(* IEC 61131-3 sources: daoli-st-library/DL_Process (part 21) *)

(* ---- FB_DL_AnnealCoolRateCtrl.st ---- *)
(*
  Name: FB_DL_AnnealCoolRateCtrl
  Category: DL_Process
  Version: 1.0.0
  Round: R89 / 2026-11-25
  开源溯源：clean-room 自研（族 锻造加热退火，ST 开源生态实测 0 命中，无外部代码引入）
  功能：退火冷却速率控制：微分实测降温速率，超速报警；同时做超温（实测高于设定 + 容差）保护。
  边界条件：① 四浮点入参全部过非有限闸；配置越域或失能进冻结分支：输出保持末值 + xValid = FALSE（R191）；
            ② 归因分离（R190）：超速与超温各有独立内部成员 _bOverRate / _bOverTemp，出口合并为 xRateAlarm，
               两成因赋值点互不共用，头注释声明合并口径；
            ③ 微分为一阶差分：速率 = (上拍温度 − 本拍温度)/周期 × 60，正值为降温方向 [℃/min]；
            ④ 首扫 _bInit 以当前温度播种上拍快照，避免首拍出现虚假大速率；非法周期取 10 ms 缺省。
  量纲自证：℃ ÷ s × 60 = ℃/min；容差 ℃ 与温度同量纲。
*)
FUNCTION_BLOCK FB_DL_AnnealCoolRateCtrl
VAR_INPUT
    xEnable : BOOL;             (* 使能 [-] Enable *)
    fTempActC : REAL;           (* 炉温实测 [℃] Furnace temperature actual [degC] *)
    fTempSpC : REAL;            (* 炉温设定 [℃] Furnace temperature setpoint [degC] *)
    fCoolRateMaxCpm : REAL;     (* 最大允许降温速率 [℃/min] Maximum allowed cooling rate [degC/min] *)
    fCycleS : REAL;             (* 扫描周期 [s] Scan cycle [s] *)
END_VAR
VAR_OUTPUT
    fRateActCpm : REAL;         (* 实测降温速率（正值为降温） [℃/min] Actual cooling rate [degC/min] *)
    xRateAlarm : BOOL;          (* 超速或超温报警（归因见内部成员） [-] Over-rate or over-temperature alarm *)
    xValid : BOOL;              (* 配置与链路有效 [-] Configuration and chain valid *)
END_VAR
VAR
    _bInit : BOOL := FALSE;     (* 首扫初始化标志 [-] First-scan init flag *)
    _bCfgBad : BOOL := FALSE;   (* 配置非法当拍量 [-] Configuration bad *)
    _bCalcOk : BOOL := FALSE;   (* 本拍计算有效 [-] Calculation valid this scan *)
    _bOverRate : BOOL := FALSE; (* 超速成因（独立成员） [-] Over-rate cause *)
    _bOverTemp : BOOL := FALSE; (* 超温成因（独立成员） [-] Over-temperature cause *)
    _fPrev : REAL := 0.0;       (* 上拍温度快照（首扫播种） [℃] Previous temperature snapshot [degC] *)
    _fRate : REAL := 0.0;       (* 速率保持量 [℃/min] Rate hold [degC/min] *)
    _fCy : REAL := 0.01;        (* 当拍有效周期 [s] Effective cycle [s] *)
END_VAR
VAR CONSTANT
    DL_ACRC_EPS : REAL := 1.0E-9;       (* 判据容差 [-] Criterion tolerance *)
    DL_ACRC_CYDEF : REAL := 0.01;       (* 缺省扫描周期 [s] Default scan cycle [s] *)
    DL_ACRC_SECMIN : REAL := 60.0;      (* 每秒 → 每分钟换算 [s/min] Second to minute *)
    DL_ACRC_TOL : REAL := 5.0;          (* 超温容差 [℃] Over-temperature tolerance [degC] *)
    DL_ACRC_TMIN : REAL := 0.0;         (* 温度下限 [℃] Temperature floor [degC] *)
    DL_ACRC_TMAX : REAL := 1400.0;      (* 温度上限 [℃] Temperature ceiling [degC] *)
    DL_ACRC_RMIN : REAL := 0.1;         (* 允许速率下限 [℃/min] Rate floor [degC/min] *)
    DL_ACRC_RMAX : REAL := 100.0;       (* 允许速率上限 [℃/min] Rate ceiling [degC/min] *)
END_VAR
(* 首扫初始化：以当前温度播种上拍快照，避免虚假大速率（R310） *)
IF NOT _bInit THEN
    _fPrev := fTempActC;
    _fRate := 0.0;
    _bInit := TRUE;
END_IF
(* 周期派生：非法周期取 10 ms 缺省（步长不塌零，除零结构性排除） *)
IF (fCycleS > 0.0) AND (fCycleS <= 1.0) THEN
    _fCy := fCycleS;
ELSE
    _fCy := DL_ACRC_CYDEF;
END_IF
(* 非有限闸（NaN 自反 + Inf 差值自减）+ 组态域闸：四浮点入参全枚举（R272） *)
_bCfgBad := (fTempActC <> fTempActC) OR ((fTempActC - fTempActC) <> 0.0)
         OR (fTempSpC <> fTempSpC) OR ((fTempSpC - fTempSpC) <> 0.0)
         OR (fCoolRateMaxCpm <> fCoolRateMaxCpm) OR ((fCoolRateMaxCpm - fCoolRateMaxCpm) <> 0.0)
         OR (fCycleS <> fCycleS) OR ((fCycleS - fCycleS) <> 0.0)
         OR (fTempActC < DL_ACRC_TMIN) OR (fTempActC > DL_ACRC_TMAX)
         OR (fTempSpC < DL_ACRC_TMIN) OR (fTempSpC > DL_ACRC_TMAX)
         OR (fCoolRateMaxCpm < DL_ACRC_RMIN) OR (fCoolRateMaxCpm > DL_ACRC_RMAX);
_bCalcOk := xEnable AND (NOT _bCfgBad);
IF _bCalcOk THEN
    (* 一阶差分：正值为降温方向，量纲 ℃/s × 60 = ℃/min *)
    _fRate := ((_fPrev - fTempActC) / _fCy) * DL_ACRC_SECMIN;
    (* 归因分离：超速与超温各写各的成员，互不共用赋值点（R190） *)
    _bOverRate := _fRate > fCoolRateMaxCpm;
    _bOverTemp := fTempActC > (fTempSpC + DL_ACRC_TOL);
    (* 快照推进放在有效计算之后，冻结时快照不动 *)
    _fPrev := fTempActC;
ELSE
    _bOverRate := FALSE;
    _bOverTemp := FALSE;
    _fPrev := fTempActC;                    (* 冻结拍也同步快照，恢复时不产生阶跃虚假速率 *)
END_IF
(* 统一出口（单点赋值）：冻结分支保持末次有效速率，保持量为已过闸的有限值（R273） *)
fRateActCpm := _fRate;
xRateAlarm := (_bOverRate OR _bOverTemp) AND _bCalcOk;
xValid := _bCalcOk;
END_FUNCTION_BLOCK

(* ---- FB_DL_BacdHvacPoll.st ---- *)
(*
  ==================================================================
  组件名 Component  : FB_DL_BacdHvacPoll
  分类   Category   : DL_Process
  版本   Version    : 1.0.1
  功能   Purpose    : BA 顺控 BACnet / Modbus 轮询行。按固定轮询间隔对 1..16 台现场
                      设备做轮询：发出轮询触发后等响应超时窗，收到响应即置在线位并
                      清重试计数；超时即重试，重试次数用尽置离线位。每轮完成后索引
                      前进并跳过离线设备（全部离线时仍逐台尝试以探测恢复），并输出
                      在线 / 离线掩码字、轮询计数与超时计数。
  溯源   Origin     : BACnet / Modbus 轮询调度为公开现场总线通信语义；本件为 clean-room
                      实现，仅借鉴来源分类与参数域组织（来源标签 roadmap-p2-bacd），
                      道莅原创设计，未复制任何闭源代码行。
  平台   Platform   : 纯 IEC 61131-3（TON / R_TRIG / WORD / SHL，无私有库）
  作者   Author     : 道莅代码库 · PLC 编程专家（R55）
  ------------------------------------------------------------------
  同拍双窗配比约束（R100）：tRespTo 必须小于 tPollInt —— 响应超时窗短于轮询间隔窗，
                      两窗职责分离：tPollInt 定节拍，tRespTo 判单台失败；超时窗覆盖整个
                      间隔会使下一拍无法发出轮询，配比反置在组态域闸内直接判故障。
  边界 Boundary     :
                      一 本件只出轮询触发与在线掩码，不做协议编解码、不写设备（属主边界）；
                      二 轮询间隔用自复位周期 TON（周期脉冲发生器用法，R328 适用方向）；
                      三 响应超时件 IN 串「等待响应相」闸与「响应已到」补集，不跨相累计；
                      四 设备索引一律回钳 1..16，跳过离线设备的循环有守护上限防死循环；
                      五 无全局变量、无外部变量声明、无物理地址寻址；
                      六 eNoDevice 为预留恒空成员：设备数为零已由组态域闸判
                         eCfgIllegal（故障级），信息级 eNoDevice 不可达，保留成员
                         以稳定接口（R56 返修留痕）。
  输出契约 Output contract:
                      nPollIdx 为当前轮询设备号（1..nDevCount），无设备时保持 1；
                      wOnlineMask / wOfflineMask 位 i-1 对应设备 i，
                      自证向量：仅 1 号设备离线 → 16#0001，仅 16 号设备离线 → 16#8000；
                      bPollTrig 与 bRespTimeout 各为单拍脉冲（内部位置位、出口映射后撤销）；
                      eCause 故障级成因与 bError 配对（R45），信息级永不置 bError。
  修订记录 Revision  :
    2026-11-20  v1.0.0  R55 首版（批 4 · 序号 20）
    2026-11-20  v1.0.1  R56 返修（7.1）：段 7 删除恒假死分支（判量 _nUseCount 经段 3
                        回钳恒 ≥1，信息级 eNoDevice 不可达），「设备数为零」语义改由
                        组态域闸 eCfgIllegal（故障级）承载；_nCurRetry 声明经核验
                        已在 VAR 区在位（7 处引用合法）。
  ==================================================================
*)

TYPE E_DL_BhdPhase :
(
    eIdle  := 0,        // 空闲：未使能或已停轮询 / idle, disabled or polling stopped
    ePoll  := 10,       // 发出：本拍发出轮询触发 / issuing, the poll trigger is raised this scan
    eWait  := 20,       // 等响应：等响应或超时 / waiting, for the response or the timeout
    eFault := 90        // 故障：组态非法锁存 / fault, illegal configuration latched
);
END_TYPE

TYPE E_DL_BhdCause :
(
    eNone       := 0,   // 无成因 / no cause
    eCfgIllegal := 1,   // 组态非法：设备数、重试上限或时间引脚越域（故障级，与 bError 配对）/ illegal config, device count, retry cap or time pin out of domain
    eDevOffline := 2,   // 有设备重试用尽转离线（信息级）/ a device exhausted its retries and went offline, informational
    eAllOffline := 3,   // 全部设备离线，仍逐台尝试探测恢复（信息级）/ every device is offline and the scan still probes for recovery
    eNoDevice   := 4    // 设备数为零（预留恒空，语义由 eCfgIllegal 承载，R56 留痕）/ no device configured, reserved always empty, carried by eCfgIllegal
);
END_TYPE

FUNCTION_BLOCK FB_DL_BacdHvacPoll
VAR_INPUT
    bEnable     : BOOL := TRUE;              // 使能，失能时停轮询并保持掩码 [-] / enable, polling stops and the masks hold when disabled
    bReset      : BOOL := FALSE;            // 复位上升沿清故障锁存、掩码与重试 [-] / reset rising edge clears the fault latch, the masks and the retries
    nDevCount   : INT := 8;                  // 轮询设备数 [台]，域 1..16 / polled device count [unit], domain 1 to 16
    nRetryMax   : INT := 2;                  // 单设备重试上限 [次]，域 0..9 / per device retry ceiling [count], domain 0 to 9
    tPollInt    : TIME := T#1S;              // 轮询间隔 [毫秒]，域 大于零 / poll interval [millisecond], domain above zero
    tRespTo     : TIME := T#500MS;           // 响应超时 [毫秒]，域 大于零 / response timeout [millisecond], domain above zero
    bRespPulse  : BOOL := FALSE;             // 响应到达脉冲（对应当前轮询设备）[-] / response arrival pulse for the currently polled device
END_VAR
VAR_OUTPUT
    nPollIdx    : INT := 1;                  // 当前轮询设备号 [设备号] / currently polled device number
    bPollTrig   : BOOL := FALSE;             // 轮询触发单拍脉冲 [-] / poll trigger single-shot pulse
    bRespTimeout: BOOL := FALSE;             // 响应超时单拍脉冲 [-] / response timeout single-shot pulse
    wOnlineMask : WORD := 16#0000;           // 在线设备掩码，位 i-1 对应设备 i [-] / online device mask, bit i minus one maps to device i
    wOfflineMask: WORD := 16#0000;           // 离线设备掩码，位 i-1 对应设备 i [-] / offline device mask, bit i minus one maps to device i
    uPollCnt    : UDINT := 0;                // 累计轮询次数（饱和到上限）[次] / total poll count, saturated [count]
    uTimeoutCnt : UDINT := 0;                // 累计响应超时次数（饱和到上限）[次] / total response timeout count, saturated [count]
    nOfflineCnt : INT := 0;                  // 当前离线设备数 [台] / current offline device count [unit]
    nCurRetry   : INT := 0;                  // 当前设备已重试次数 [次] / retries already spent on the current device [count]
    ePhase      : E_DL_BhdPhase := E_DL_BhdPhase.eIdle; // 相位出口 [枚举] / phase outlet [enum]
    eCause      : E_DL_BhdCause := E_DL_BhdCause.eNone; // 成因出口 [枚举] / cause outlet [enum]
    bError      : BOOL := FALSE;             // 故障锁存标志 [-] / fault latch flag
END_VAR
VAR
    rtResp      : R_TRIG;                    // 响应沿检测，段 0 无条件刷新 / response edge detector, refreshed unconditionally in segment zero
    rtReset     : R_TRIG;                    // 复位沿检测，段 0 无条件刷新 / reset edge detector, refreshed unconditionally in segment zero
    tonPollInt  : TON;                       // 轮询间隔周期计时（自复位式）/ poll interval timer, self resetting
    tonResp     : TON;                       // 响应超时计时，段 0 无条件刷新 / response timeout timer, refreshed unconditionally in segment zero
    _ePhase     : E_DL_BhdPhase := E_DL_BhdPhase.eIdle;   // 内部相位，CASE 唯一写入目标 / internal phase, the only CASE write target
    _eCause     : E_DL_BhdCause := E_DL_BhdCause.eNone;   // 信息级成因，每拍重算 / informational cause, recomputed every scan
    _eFaultCause: E_DL_BhdCause := E_DL_BhdCause.eNone;   // 故障级成因，锁存至复位沿 / fault cause, latched until the reset edge
    _bFault     : BOOL := FALSE;             // 故障锁存位 [-] / fault latch bit
    _bInit      : BOOL := FALSE;             // 首扫初始化完成标志（R310）/ first scan initialisation flag
    _bCfgBad    : BOOL := FALSE;             // 组态非法判定 [-] / illegal configuration verdict
    _bPollInt   : BOOL := FALSE;             // 轮询触发内部位，统一出口映射 / internal poll trigger bit, mapped at the unified outlet
    _bToInt     : BOOL := FALSE;             // 超时脉冲内部位，统一出口映射 / internal timeout bit, mapped at the unified outlet
    _bOfflineNew: BOOL := FALSE;             // 本拍有新设备转离线 [-] / a device went offline this scan
    _bAllOff    : BOOL := FALSE;             // 全部设备离线 [-] / every device is offline
    _bFound     : BOOL := FALSE;             // 跳过循环命中标志 [-] / hit flag of the skip loop
    _bIsOffline : BOOL := FALSE;             // 被检设备是否离线 [-] / whether the checked device is offline
    _nUseCount  : INT := 1;                  // 钳定后的设备数 [台] / clamped device count [unit]
    _nRetryUse  : INT := 1;                  // 钳定后的重试上限 [次] / clamped retry ceiling [count]
    _nIdx       : INT := 1;                  // 设备索引（回钳 1..16）[设备号] / device index clamped one through sixteen
    _nGuard     : INT := 0;                  // 跳过循环守护计数 [次] / skip loop guard [count]
    _nIdxProbe  : INT := 1;                  // 离线统计探测索引 [设备号] / probe index for the offline statistics
    _nCurRetry  : INT := 0;                  // 当前设备重试计数（声明补齐，R55 终审）/ current device retry counter, declaration completed at R55 review
    _nOfflineCnt: INT := 0;                  // 本轮统计离线设备数工作值（出口映射源）[台] / offline device count working value, source of the outlet [unit]
    _wOff       : WORD := 16#0000;           // 离线掩码工作字 / offline mask working word
    _wOn        : WORD := 16#0000;           // 在线掩码工作字（按位或累计）/ online mask working word
    _wBit       : WORD := 16#0001;           // 本设备位掩码，先移位后置位（R327）/ device bit mask, shift before setting
    _uPoll      : UDINT := 0;                // 轮询计数工作值 [次] / poll count working value [count]
    _uTo        : UDINT := 0;                // 超时计数工作值 [次] / timeout count working value [count]
END_VAR
VAR CONSTANT
    DL_BHD_MAX      : INT := 16;             // 设备容量与索引回钳上界 [台] / device capacity and index clamp upper bound
    DL_BHD_RETRY_MAX: INT := 9;              // 重试上限的钳定上限 [次] / clamp ceiling of the retry cap [count]
    DL_BHD_CNT_MAX  : UDINT := 2000000000;   // 计数饱和上限（常量在 DINT 可表范围内）[次] / count saturation ceiling, the constant fits in DINT
    DL_BHD_MASK_NONE: WORD := 16#0000;       // 空掩码常量 [-] / empty mask constant
    DL_BHD_MASK_ONE : WORD := 16#0001;       // 单位位常量 [-] / single bit constant
END_VAR

// 段 0｜定时器与沿检测无条件周期刷新（禁入分支）；轮询间隔用自复位式周期发生器 / segment 0, unconditional refresh with a self resetting periodic generator
rtResp(CLK := bRespPulse); // 响应沿无条件刷新 / unconditional refresh of the response edge
rtReset(CLK := bReset); // 复位沿无条件刷新 / unconditional refresh of the reset edge
tonPollInt(IN := (NOT tonPollInt.Q) AND bEnable AND (NOT _bFault), PT := tPollInt); // 轮询间隔周期发生器，Q 到时下一拍即重启（R328 周期脉冲方向）/ periodic poll generator that restarts right after its own pulse
tonResp(IN := (_ePhase = E_DL_BhdPhase.eWait) AND (NOT rtResp.Q) AND (NOT _bFault), PT := tRespTo); // 响应超时，IN 串等待相闸与响应到达补集 / response timeout with the waiting gate and the response complement on IN

// 段 1｜首扫初始化（R310）/ segment 1, first scan initialisation
IF NOT _bInit THEN // 首扫一拍 / the very first scan
    _bInit := TRUE; // 置首扫完成标志 / raise the first scan flag
    _ePhase := E_DL_BhdPhase.eIdle; // 相位从空闲起步 / the phase starts from idle
    _eCause := E_DL_BhdCause.eNone; // 信息级成因清零 / clear the informational cause
    _eFaultCause := E_DL_BhdCause.eNone; // 故障级成因清零 / clear the fault cause
    _bFault := FALSE; // 故障锁存清零 / clear the fault latch
    _wOff := DL_BHD_MASK_NONE; // 离线掩码清零 / clear the offline mask
    _wOn := DL_BHD_MASK_NONE; // 在线掩码清零 / clear the online mask
    _nIdx := 1; // 索引归位 / park the index at one
    _uPoll := 0; // 轮询计数清零 / clear the poll count
    _uTo := 0; // 超时计数清零 / clear the timeout count
END_IF

// 段 2｜复位沿作用域：清锁存 / 清掩码 / 清计数与索引（四项逐项声明）/ segment 2, reset edge scope declared item by item
IF rtReset.Q THEN // 复位沿 / reset edge
    _bFault := FALSE; // 作用域一：清故障锁存 / scope one, clear the fault latch
    _eFaultCause := E_DL_BhdCause.eNone; // 作用域一：清故障级成因 / scope one, clear the fault cause
    _wOff := DL_BHD_MASK_NONE; // 作用域二：清离线掩码 / scope two, clear the offline mask
    _wOn := DL_BHD_MASK_NONE; // 作用域二：清在线掩码 / scope two, clear the online mask
    _nIdx := 1; // 作用域三：索引归位 / scope three, park the index
    _nCurRetry := 0; // 作用域三：清重试计数 / scope three, clear the retry count
    _ePhase := E_DL_BhdPhase.eIdle; // 作用域四：迁回空闲相 / scope four, migrate back to idle
    _bPollInt := FALSE; // 作用域四：清轮询脉冲内部位 / scope four, clear the internal poll bit
    _bToInt := FALSE; // 作用域四：清超时脉冲内部位 / scope four, clear the internal timeout bit
END_IF

// 段 3｜组态域闸（R151 全覆盖）/ segment 3, configuration domain gate over every pin
_bCfgBad := FALSE; // 组态非法预置假 / preset the illegal configuration verdict to false
IF (nDevCount < 1) OR (nDevCount > DL_BHD_MAX) THEN // 设备数越域 / the device count is out of domain
    _bCfgBad := TRUE; // 判非法 / mark illegal
END_IF
IF (nRetryMax < 0) OR (nRetryMax > DL_BHD_RETRY_MAX) THEN // 重试上限越域 / the retry cap is out of domain
    _bCfgBad := TRUE; // 判非法 / mark illegal
END_IF
IF (tPollInt <= T#0S) OR (tRespTo <= T#0S) THEN // 时间引脚非正 / a time pin is not positive
    _bCfgBad := TRUE; // 判非法 / mark illegal
END_IF
IF tRespTo >= tPollInt THEN // 响应超时窗不得覆盖整个轮询间隔（配比约束，R100）/ the response window must not swallow the whole poll interval
    _bCfgBad := TRUE; // 判非法 / mark illegal
END_IF
IF _bCfgBad AND (NOT _bFault) THEN // 组态非法且未锁存 / illegal configuration and not yet latched
    _bFault := TRUE; // 置故障锁存 / raise the fault latch
    _eFaultCause := E_DL_BhdCause.eCfgIllegal; // 故障级成因 (R45 配对 bError) / fault grade cause paired with bError
    _ePhase := E_DL_BhdPhase.eFault; // 迁故障相 / migrate to the fault phase
END_IF
_nUseCount := nDevCount; // 设备数直通 / the device count passes through
IF _nUseCount < 1 THEN // 下越界 / below the lower bound
    _nUseCount := 1; // 回钳到 1 / clamp to one
ELSIF _nUseCount > DL_BHD_MAX THEN // 上越界 / above the upper bound
    _nUseCount := DL_BHD_MAX; // 回钳到 16 / clamp to sixteen
END_IF
_nRetryUse := nRetryMax; // 重试上限直通 / the retry cap passes through
IF _nRetryUse < 0 THEN // 下越界（防御）/ below the lower bound as a defence
    _nRetryUse := 0; // 回钳到 0 / clamp to zero
ELSIF _nRetryUse > DL_BHD_RETRY_MAX THEN // 上越界 / above the upper bound
    _nRetryUse := DL_BHD_RETRY_MAX; // 回钳到 9 / clamp to nine
END_IF
IF _nIdx < 1 THEN // 索引下越界 / the index is below the lower bound
    _nIdx := 1; // 回钳到 1 / clamp to one
ELSIF _nIdx > _nUseCount THEN // 索引上越界 / the index is above the upper bound
    _nIdx := _nUseCount; // 回钳到末台 / clamp to the last unit
END_IF

// 段 4｜失效使能与设备位更新 / segment 4, enable handling and device bit updates
_eCause := E_DL_BhdCause.eNone; // 信息级成因每拍重算 / the informational cause is recomputed every scan
_bOfflineNew := FALSE; // 新转离线标志预置假 / preset the new offline flag to false
_bAllOff := FALSE; // 全离线标志每拍重算 / the all offline flag is recomputed every scan
IF NOT bEnable THEN // 失能：停轮询并保持掩码（R191 显式声明）/ disabled, polling stops and the masks hold
    _ePhase := E_DL_BhdPhase.eIdle; // 回空闲相 / return to idle
    _bPollInt := FALSE; // 撤轮询脉冲内部位 / withdraw the internal poll bit
    _bToInt := FALSE; // 撤超时脉冲内部位 / withdraw the internal timeout bit
END_IF
_wBit := SHL(DL_BHD_MASK_ONE, _nIdx - 1); // 当前设备位掩码，位移量 0..15 由索引回钳与容量常量证明 / the current device bit mask, the shift zero through fifteen is proven by the index clamp and the capacity constant
IF rtResp.Q AND (_ePhase = E_DL_BhdPhase.eWait) THEN // 等待相收到响应 / a response arrived while waiting
    _wOff := _wOff AND NOT _wBit; // 清离线位 / clear the offline bit
    _wOn := _wOn OR _wBit; // 置在线位 / set the online bit
    _nCurRetry := 0; // 清重试计数 / clear the retry count
    _ePhase := E_DL_BhdPhase.ePoll; // 本轮结束，转下一轮发出相 / the round is finished and the next issuing phase follows
    _bFound := FALSE; // 跳过命中标志预置假 / preset the skip hit flag to false
    _nGuard := 0; // 守护计数清零 / reset the guard
    WHILE (_nGuard < DL_BHD_MAX) AND (NOT _bFound) DO // 跳过离线设备，守护上限为容量 / skip offline devices with the capacity as the guard
        _nGuard := _nGuard + 1; // 守护计数递增 / increment the guard
        _nIdx := _nIdx + 1; // 索引前进 / advance the index
        IF _nIdx > _nUseCount THEN // 越过末台 / past the last unit
            _nIdx := 1; // 回卷到首台 / wrap back to the first unit
        END_IF
        _wBit := SHL(DL_BHD_MASK_ONE, _nIdx - 1); // 候选设备位掩码 / the candidate device bit mask
        _bIsOffline := ((_wOff AND _wBit) <> DL_BHD_MASK_NONE); // 候选设备是否离线 / whether the candidate is offline
        IF NOT _bIsOffline THEN // 候选在线 / the candidate is online
            _bFound := TRUE; // 命中 / hit
        END_IF
    END_WHILE
    IF NOT _bFound THEN // 全部离线，仍逐台尝试（探测恢复）/ every device is offline and probing continues
        _nIdx := _nIdx + 1; // 索引照常前进 / the index advances anyway
        IF _nIdx > _nUseCount THEN // 越过末台 / past the last unit
            _nIdx := 1; // 回卷到首台 / wrap back to the first unit
        END_IF
        _bAllOff := TRUE; // 置全离线标志 / raise the all offline flag
    END_IF
END_IF
IF tonResp.Q AND (_ePhase = E_DL_BhdPhase.eWait) THEN // 等待相超时 / the waiting phase timed out
    _bToInt := TRUE; // 超时脉冲内部位置位（统一出口映射，R187）/ raise the internal timeout bit, mapped at the unified outlet
    IF _uTo < DL_BHD_CNT_MAX THEN // 未达饱和上限 / below the ceiling
        _uTo := _uTo + 1; // 超时计数递增 / increment the timeout count
    END_IF
    IF _nCurRetry < _nRetryUse THEN // 重试未用尽 / retries remain
        _nCurRetry := _nCurRetry + 1; // 重试计数递增并立即重发 / increment the retry count and re-issue at once
        _ePhase := E_DL_BhdPhase.ePoll; // 回发出相重试同一台 / back to the issuing phase for the same unit
    ELSE // 重试用尽 / retries exhausted
        _wOff := _wOff OR _wBit; // 置离线位 / set the offline bit
        _wOn := _wOn AND NOT _wBit; // 清在线位 / clear the online bit
        _bOfflineNew := TRUE; // 记新转离线 / record the new offline event
        _nCurRetry := 0; // 重试计数清零 / clear the retry count
        _ePhase := E_DL_BhdPhase.ePoll; // 回发出相转下一台 / back to the issuing phase for the next unit
        _bFound := FALSE; // 跳过命中标志预置假 / preset the skip hit flag to false
        _nGuard := 0; // 守护计数清零 / reset the guard
        WHILE (_nGuard < DL_BHD_MAX) AND (NOT _bFound) DO // 跳过离线设备 / skip offline devices
            _nGuard := _nGuard + 1; // 守护计数递增 / increment the guard
            _nIdx := _nIdx + 1; // 索引前进 / advance the index
            IF _nIdx > _nUseCount THEN // 越过末台 / past the last unit
                _nIdx := 1; // 回卷到首台 / wrap back to the first unit
            END_IF
            _wBit := SHL(DL_BHD_MASK_ONE, _nIdx - 1); // 候选设备位掩码 / the candidate device bit mask
            _bIsOffline := ((_wOff AND _wBit) <> DL_BHD_MASK_NONE); // 候选设备是否离线 / whether the candidate is offline
            IF NOT _bIsOffline THEN // 候选在线 / the candidate is online
                _bFound := TRUE; // 命中 / hit
            END_IF
        END_WHILE
        IF NOT _bFound THEN // 全部离线 / every device is offline
            _bAllOff := TRUE; // 置全离线标志 / raise the all offline flag
        END_IF
    END_IF
END_IF

// 段 5｜相位机：ENUM + CASE，含 ELSE 非法相位兜底（R128）/ segment 5, phase machine with an ELSE fallback for illegal phases
CASE _ePhase OF
E_DL_BhdPhase.eIdle: // 空闲相：使能且无故障才起轮询 / idle, polling starts when enabled and unfaulted
    IF bEnable AND (NOT _bFault) THEN // 使能且无故障 / enabled and unfaulted
        _ePhase := E_DL_BhdPhase.ePoll; // 迁发出相 / migrate to the issuing phase
    END_IF

E_DL_BhdPhase.ePoll: // 发出相：本拍发轮询触发并转等待相 / issuing phase, the trigger is raised and the waiting phase follows
    IF bEnable AND (NOT _bFault) AND tonPollInt.Q THEN // 轮询间隔到 / the poll interval elapsed
        _bPollInt := TRUE; // 轮询触发内部位置位（统一出口映射，R187）/ raise the internal poll bit, mapped at the unified outlet
        IF _uPoll < DL_BHD_CNT_MAX THEN // 未达饱和上限 / below the ceiling
            _uPoll := _uPoll + 1; // 轮询计数递增 / increment the poll count
        END_IF
        _ePhase := E_DL_BhdPhase.eWait; // 迁等待相 / migrate to the waiting phase
    END_IF

E_DL_BhdPhase.eWait: // 等待相：等响应或超时（两出口均在段 4 处理）/ waiting phase, the response and the timeout are handled in segment four
    IF (NOT bEnable) OR _bFault THEN // 失能或故障 / disabled or faulted
        _ePhase := E_DL_BhdPhase.eIdle; // 回空闲相 / return to idle
    END_IF

E_DL_BhdPhase.eFault: // 故障相：停轮询，等复位沿 / fault phase, polling stopped until the reset edge
    _bPollInt := FALSE; // 撤轮询脉冲内部位 / withdraw the internal poll bit
    _bToInt := FALSE; // 撤超时脉冲内部位 / withdraw the internal timeout bit
    _nCurRetry := 0; // 清重试计数 / clear the retry count

ELSE // 非法相位兜底（R128）/ illegal phase fallback
    _bFault := TRUE; // 置故障锁存 / raise the fault latch
    _eFaultCause := E_DL_BhdCause.eCfgIllegal; // 故障级成因记组态非法 / record the illegal configuration cause
    _ePhase := E_DL_BhdPhase.eFault; // 迁故障相 / migrate to the fault phase
END_CASE

// 段 6｜离线统计：逐台扫全容量统计，未参与设备按零位计 / segment 6, offline statistics over the full capacity
_nOfflineCnt := 0; // 离线计数清零 / clear the offline count
_nIdxProbe := 1; // 探测索引自 1 起 / the probe index starts at one
WHILE _nIdxProbe <= DL_BHD_MAX DO // 全容量扫查，未参与设备恒为零位 / sweep the full capacity because unused devices stay cleared
    _wBit := SHL(DL_BHD_MASK_ONE, _nIdxProbe - 1); // 本设备位掩码 / this device bit mask
    IF ((_wOff AND _wBit) <> DL_BHD_MASK_NONE) THEN // 本设备离线 / this device is offline
        _nOfflineCnt := _nOfflineCnt + 1; // 离线计数递增 / increment the offline count
    END_IF
    _nIdxProbe := _nIdxProbe + 1; // 索引递增 / increment the index
END_WHILE

// 段 7｜成因分派（固定优先级：故障 > 新转离线 > 全离线 > 无设备 > 无成因）/ segment 7, cause dispatch with a fixed priority
IF _bFault THEN // 故障锁存优先 / the fault latch takes priority
    eCause := _eFaultCause; // 故障级成因锁存回放 / the fault cause is replayed from the latch
ELSIF _bOfflineNew THEN // 本拍有新设备转离线 / a device went offline this scan
    eCause := E_DL_BhdCause.eDevOffline; // 信息级成因 / informational cause
ELSIF _bAllOff THEN // 全部离线 / every device is offline
    eCause := E_DL_BhdCause.eAllOffline; // 信息级成因 / informational cause
ELSE // 设备数为零的情形已由组态域闸 eCfgIllegal 承载（R56 死分支删除留痕）/ the no device case is carried by the configuration gate
    eCause := _eCause; // 信息级成因直映 / the informational cause is mapped directly
END_IF

// 段 8｜统一出口 / segment 8, unified outlet
nPollIdx := _nIdx; // 当前轮询设备号出口 / currently polled device outlet
bPollTrig := _bPollInt; // 轮询触发映射本拍值 / map the poll trigger for this scan
_bPollInt := FALSE; // 映射后立即撤销，保证单拍宽度（R187 两段式）/ revoke right after mapping to keep a single-scan width
bRespTimeout := _bToInt; // 超时脉冲映射本拍值 / map the timeout pulse for this scan
_bToInt := FALSE; // 映射后立即撤销，保证单拍宽度（R187 两段式）/ revoke right after mapping to keep a single-scan width
wOnlineMask := _wOn; // 在线掩码出口 / online mask outlet
wOfflineMask := _wOff; // 离线掩码出口 / offline mask outlet
uPollCnt := _uPoll; // 轮询计数出口 / poll count outlet
uTimeoutCnt := _uTo; // 超时计数出口 / timeout count outlet
nOfflineCnt := _nOfflineCnt; // 离线设备数出口 / offline device count outlet
nCurRetry := _nCurRetry; // 当前重试次数出口 / current retry count outlet
ePhase := _ePhase; // 相位出口单点映射 / single-point phase outlet mapping
bError := _bFault; // 故障标志与锁存位同源 / the fault flag shares the latch source
END_FUNCTION_BLOCK

(* ---- FB_DL_BatchDeviationAlarm.st ---- *)
//==============================================================================
// 功能块：FB_DL_BatchDeviationAlarm ｜ 中文名称：批次偏差分级报警与首出归因
// 所属子库：DL_Process ｜ 版本：v1.0.0 ｜ 兼容：CODESYS V3.5+ / TwinCAT 3 / 汇川 InoProShop
// 功能描述：批次偏差四档分级监视——|测量 - 设定| 越档判定：预警档
//           （fBandWarn < |偏差| <= fBandMinor）、次要档（<= fBandMajor）、
//           严重档（> fBandMajor），越限须持续 tDebounce 才确认（防瞬时
//           噪声）；首出归因：首个非正常档确认时锁存档位与方向（高/低
//           向），锁存至 bReset，后续档位波动不重写首因（归因证据链，
//           R81 还原方向不饱和同理）。严重档确认为故障级（置 bError），
//           预警/次要档为信息级。
// 开源溯源 (Origin)：道莅原创实现（参考批次过程偏差分级与首出报警（first-out）工程惯例 分类与参数域）
// 单位表：偏差[工艺量纲（与 fValueMeas/fValueSp 同量纲）] / 带宽[同量纲] /
//         时间[ms]
// 错误码表：16#0005_01FA 信息级（预警/次要档偏差激活确认，不置 bError）/
//           16#0005_01FB 信息级（首出归因锁存已建立，不置 bError）/
//           16#0005_033C 故障级（组态非法：带宽非单调（须 0 < 预警 <
//           次要 < 严重）或任一输入非有限，置 bError）/ 16#0005_033D
//           故障级（严重档偏差确认：去抖后仍 > fBandMajor，置 bError，
//           并建立首出锁存——该场景不可由 033C 的组态类判据观测，属
//           工艺偏差独立域）/ 16#0005_033E 故障级兜底（状态机落 ELSE，
//           置 bError）
// 状态机：E_DL_BatchDevState（四态：eIdle=0 / eMonitor=10 / eFault=99，
//           外加 eDeviated=20 激活保持态），CASE 含 ELSE 兜底，ELSE 置
//           033E 并输出正常档
// 边界行为：① 组态非法 → 故障态锁存，bReset 复位；② 越限去抖未满判据
//           消失 → 不确认（防瞬时噪声）；③ 偏差回落至正常带 → 回监视
//           态（首出锁存保持，bReset 才清）；④ 首出锁存仅在无锁存时
//           建立（首出语义，后续波动不重写）；⑤ 未使能输出正常档且
//           bValid := FALSE；⑥ 安全侧 = 故障路径偏差档位输出严重档
//           （不可信数据按最坏档呈现）。
// 修订历史：v1.0.0 2026-11-17 首版（R24 派单 · ROADMAP P1 §734）
//==============================================================================

(*------------------------------------------------------------------------------
 * 枚举: E_DL_BatchDevLevel（归属本功能块，同文件发布，全库唯一定义）
 * 含义: 偏差四档分级（档位 0..3，对应越限带宽递增）。
 *-----------------------------------------------------------------------------*)
TYPE E_DL_BatchDevLevel :
(
    eNormal := 0,   // 正常：偏差在预警带内 / Normal, deviation inside the warn band
    eWarn   := 1,   // 预警：|偏差| > 预警带 / Warn, deviation beyond the warn band
    eMinor  := 2,   // 次要：|偏差| > 次要带 / Minor, deviation beyond the minor band
    eMajor  := 3    // 严重：|偏差| > 严重带（故障级） / Major, deviation beyond the major band, fault class
);
END_TYPE

(*------------------------------------------------------------------------------
 * 枚举: E_DL_BatchDevState（归属本功能块，同文件发布，全库唯一定义）
 * 含义: 分级监视相位，每个成员在 CASE 中有且仅有一个标签。
 *-----------------------------------------------------------------------------*)
TYPE E_DL_BatchDevState :
(
    eIdle     := 0,   // 空闲：未使能 / Idle, not enabled
    eMonitor  := 10,  // 监视：档位判定与去抖 / Monitor, level verdict and debounce
    eDeviated := 20,  // 激活保持：非正常档确认保持 / Deviated, non-normal level held
    eFault    := 99   // 故障：组态非法/非法状态 / Fault, config or illegal state
);
END_TYPE

FUNCTION_BLOCK FB_DL_BatchDeviationAlarm
VAR_INPUT
    bEnable     : BOOL;                     // 分级监视使能 [—] / Monitoring enable
    bReset      : BOOL;                     // 故障/首出复位 [—]，上升沿清首出锁存 / Fault and first-out reset, rising edge clears latches
    fValueMeas  : LREAL;                    // 批次实测值 [工艺量纲] / Batch measured value [process unit]
    fValueSp    : LREAL;                    // 批次设定值 [工艺量纲] / Batch setpoint [process unit]
    fBandWarn   : LREAL := 1.0;             // 预警带宽 [工艺量纲]，须 > 0 / Warn band width [process unit]
    fBandMinor  : LREAL := 2.0;             // 次要带宽 [工艺量纲]，须 > 预警带宽 / Minor band width [process unit]
    fBandMajor  : LREAL := 5.0;             // 严重带宽 [工艺量纲]，须 > 次要带宽 / Major band width [process unit]
    tDebounce   : TIME  := T#2S;            // 越限去抖窗 [ms]，须 > 0 / Violation debounce window [ms]
END_VAR
VAR_OUTPUT
    eDevLevel    : E_DL_BatchDevLevel;      // 当前偏差档位 [—] / Current deviation level
    fDeviation   : LREAL;                   // 当前偏差 [工艺量纲]（带符号，诊断出口） / Current deviation [process unit], signed, diagnostics
    bFirstOut    : BOOL;                    // 首出锁存有效 [—]（bReset 才清） / First-out latch valid, cleared by reset
    eFirstOut    : E_DL_BatchDevLevel;      // 首出档位 [—] / First-out level
    bFirstHigh   : BOOL;                    // 首出方向 [—]，TRUE = 高向 / First-out direction, TRUE high side
    eState       : E_DL_BatchDevState;      // 相位出口 [—] / Phase outlet
    eErr         : UDINT;                   // 错误码，0 = 无错，码位 16#0005_01FA 起信息级、16#0005_033C 起故障级（分带见错误码表） / Error code, 0 = no error, band info/fault per the code table
    bError       : BOOL;                    // 故障级标志，仅故障级错误置位 / Fault-class flag, set only on fault-level codes
    bValid       : BOOL;                    // 输出可用标志 / Outputs usable flag
END_VAR
VAR
    fbDebounce : TON;                       // 越限去抖计时（每拍无条件刷新）[ms] / Debounce timer, refreshed unconditionally
    _eState    : E_DL_BatchDevState := E_DL_BatchDevState.eIdle; // 当前相位 / Current phase
    _bCfgBad   : BOOL;                      // 组态非法锁存 / Illegal config latch
    _eLevelNow : E_DL_BatchDevLevel := E_DL_BatchDevLevel.eNormal; // 本拍档位判定 / Level verdict of this scan
    _bViolate  : BOOL;                      // 越限电平（非正常档判定） / Violation level
    _bInfoAct  : BOOL;                      // 预警/次要激活信息当拍标志 / Warn or minor activation info flag
    _bInfoFirst: BOOL;                      // 首出建立信息当拍标志 / First-out-established info flag
    _bIllegal  : BOOL;                      // 非法状态标志 / Illegal state flag
    _bInit     : BOOL := FALSE;             // 首扫标志，初值 FALSE 取非判定 / First-scan flag, tested negated
END_VAR
VAR CONSTANT
    DL_BDA_INF  : LREAL := 1.7976931348623157E308; // LREAL 幅值上限 / LREAL magnitude ceiling
    DL_BDA_EPS  : LREAL := 1.0E-6;          // 浮点判零容差 [工艺量纲] / Float zero tolerance [process unit]
    DL_BDA_ZERO : LREAL := 0.0;             // 零值常量，避免裸字面量 [混合] / Zero constant, avoids a bare literal
END_VAR

(*------------------------------------------------------------------------------
 * 段 1｜每拍预置：档位出口正常档起步（安全侧），单拍标志预清零
 *      Level outlet starts at normal, fail-safe, one-shot flags pre-cleared
 *-----------------------------------------------------------------------------*)
eDevLevel  := E_DL_BatchDevLevel.eNormal; // 档位出口先置正常（激活态在段 5 重置） / Level preset normal
fDeviation := DL_BDA_ZERO;               // 偏差出口每拍重算 / Deviation outlet recomputed
eErr   := 16#0000_0000;                  // 错误码每拍重算 / Error code recomputed
bError := FALSE;                         // 故障标志每拍重算 / Fault flag recomputed
bValid := FALSE;                         // 可用标志每拍重算 / Usable flag recomputed
_bInfoAct  := FALSE;                     // 激活信息预清零 / Activation info pre-cleared
_bInfoFirst := FALSE;                    // 首出信息预清零 / First-out info pre-cleared
_bIllegal   := FALSE;                    // 非法状态预清零 / Illegal flag pre-cleared

(*------------------------------------------------------------------------------
 * 段 2｜首扫初始化
 *      First-scan initialisation
 *-----------------------------------------------------------------------------*)
IF NOT _bInit THEN
    _eState  := E_DL_BatchDevState.eIdle; // 相位空闲起步 / Phase starts idle
    _bCfgBad := FALSE;                   // 组态锁存清零 / Config latch cleared
    bFirstOut := FALSE;                  // 首出锁存清零 / First-out latch cleared
    eFirstOut := E_DL_BatchDevLevel.eNormal; // 首出档位清零 / First-out level reset
    bFirstHigh := FALSE;                 // 首出方向清零 / First-out direction reset
    _bInit   := TRUE;                    // 首扫只做一次 / The first scan runs once
END_IF

(*------------------------------------------------------------------------------
 * 段 3｜组态防御闸：非有限（R79）+ 带宽单调域（0 < 预警 < 次要 < 严重）
 *      Configuration defense gates with the band monotonicity rule
 *-----------------------------------------------------------------------------*)
IF (fValueMeas <> fValueMeas) OR (ABS(fValueMeas) > DL_BDA_INF)
   OR (fValueSp <> fValueSp) OR (ABS(fValueSp) > DL_BDA_INF)
   OR (fBandWarn <> fBandWarn) OR (ABS(fBandWarn) > DL_BDA_INF)
   OR (fBandMinor <> fBandMinor) OR (ABS(fBandMinor) > DL_BDA_INF)
   OR (fBandMajor <> fBandMajor) OR (ABS(fBandMajor) > DL_BDA_INF) THEN
    _bCfgBad := TRUE;                    // 非有限归组态非法锁存 / Non-finite folded into the config latch
END_IF
IF (NOT _bCfgBad) AND ((fBandWarn <= DL_BDA_EPS) OR (fBandMinor <= fBandWarn)
   OR (fBandMajor <= fBandMinor) OR (tDebounce <= T#0MS)) THEN
    _bCfgBad := TRUE;                    // 带宽非单调或去抖窗非法锁存 / Non-monotonic bands or illegal window latched
END_IF
IF bReset THEN
    _bCfgBad := FALSE;                   // 复位清组态锁存 / Reset clears the config latch
    bFirstOut := FALSE;                  // 复位清首出锁存（归因证据链重开） / Reset clears the first-out latch
    eFirstOut := E_DL_BatchDevLevel.eNormal; // 复位清首出档位 / Reset clears the first-out level
    bFirstHigh := FALSE;                 // 复位清首出方向 / Reset clears the direction
END_IF

(*------------------------------------------------------------------------------
 * 段 4｜档位判定与去抖计时无条件刷新（R40：CASE 之外每拍必调）
 *      Level verdict and debounce timer refreshed unconditionally
 *-----------------------------------------------------------------------------*)
IF (NOT _bCfgBad) AND ((fValueMeas <> fValueMeas) OR (ABS(fValueMeas) > DL_BDA_INF)
   OR (fValueSp <> fValueSp) OR (ABS(fValueSp) > DL_BDA_INF)) THEN
    _eLevelNow := E_DL_BatchDevLevel.eMajor; // 运行中数据非有限按最坏档呈现（R90：033D 域复用） / Non-finite data presented as the worst level
ELSE
    fDeviation := fValueMeas - fValueSp; // 带符号偏差 [工艺量纲] / Signed deviation
    IF ABS(fDeviation) > fBandMajor THEN
        _eLevelNow := E_DL_BatchDevLevel.eMajor; // 严重档 / Major
    ELSIF ABS(fDeviation) > fBandMinor THEN
        _eLevelNow := E_DL_BatchDevLevel.eMinor; // 次要档 / Minor
    ELSIF ABS(fDeviation) > fBandWarn THEN
        _eLevelNow := E_DL_BatchDevLevel.eWarn; // 预警档 / Warn
    ELSE
        _eLevelNow := E_DL_BatchDevLevel.eNormal; // 正常档 / Normal
    END_IF
END_IF
_bViolate := (_eLevelNow <> E_DL_BatchDevLevel.eNormal); // 越限电平（任一非正常档） / Violation level
fbDebounce(IN := (_eState = E_DL_BatchDevState.eMonitor) AND _bViolate
             AND (_eLevelNow = eDevLevel), PT := tDebounce); // 越限去抖窗（同档驻留） / Debounce window on the same level

(*------------------------------------------------------------------------------
 * 段 5｜相位机（CASE 含 ELSE 兜底；状态改写只出现在分支判据内，R39）
 *      Phase machine with ELSE fallback
 *-----------------------------------------------------------------------------*)
CASE _eState OF

    E_DL_BatchDevState.eIdle:              // 空闲：使能且组态合法进监视
        IF bEnable AND (NOT _bCfgBad) THEN
            _eState := E_DL_BatchDevState.eMonitor; // 进监视 / To monitor
        ELSIF bEnable AND _bCfgBad THEN
            _eState := E_DL_BatchDevState.eFault; // 组态非法进故障 / Illegal config to fault
        END_IF

    E_DL_BatchDevState.eMonitor:           // 监视：同档越限去抖满进激活保持
        IF (NOT bEnable) OR _bCfgBad THEN
            _eState := E_DL_BatchDevState.eFault; // 异常转故障 / Anomaly, fault
        ELSIF fbDebounce.Q THEN
            IF (NOT bFirstOut) THEN
                bFirstOut := TRUE;         // 首出锁存建立（后续波动不重写，R81） / First-out latch established, never rewritten
                eFirstOut := _eLevelNow;   // 首出档位锁定 / First-out level locked
                bFirstHigh := fDeviation > DL_BDA_ZERO; // 首出方向锁定 / First-out direction locked
                _bInfoFirst := TRUE;       // 首出建立提示（信息级，拍 N 进入） / First-out notice, info
            END_IF
            IF _eLevelNow = E_DL_BatchDevLevel.eMajor THEN
                _eState := E_DL_BatchDevState.eDeviated; // 严重档确认进激活保持（故障级在段 6 报） / Major confirmed, to deviated
            ELSE
                _bInfoAct := TRUE;         // 预警/次要档激活（信息级） / Warn or minor activation, info
                _eState := E_DL_BatchDevState.eDeviated; // 进激活保持 / To deviated
            END_IF
        END_IF

    E_DL_BatchDevState.eDeviated:          // 激活保持：偏差回正常带回监视（首出锁存保持）
        IF (NOT bEnable) OR _bCfgBad THEN
            _eState := E_DL_BatchDevState.eFault; // 异常转故障 / Anomaly, fault
        ELSIF _eLevelNow = E_DL_BatchDevLevel.eNormal THEN
            _eState := E_DL_BatchDevState.eMonitor; // 回监视（首出锁存保持） / Back to monitor, first-out held
        END_IF

    E_DL_BatchDevState.eFault:             // 故障：复位沿且组态恢复回监视
        IF bReset AND (NOT _bCfgBad) THEN
            _eState := E_DL_BatchDevState.eMonitor; // 回监视 / Back to monitor
        END_IF

    ELSE                                   // 非法状态兜底（R21：CASE 必带 ELSE）
        _bIllegal := TRUE;                 // 标记非法状态 / Flag the illegal state
        eDevLevel := E_DL_BatchDevLevel.eMajor; // 最坏档呈现（安全侧） / Worst level presented
        _eState := E_DL_BatchDevState.eFault; // 回故障态 / Back to fault
END_CASE

(*------------------------------------------------------------------------------
 * 段 6｜码位出口与放行（故障级码 3 行内置 bError，R45/R101 配对）
 *      Code outlet and release, fault codes paired with bError
 *-----------------------------------------------------------------------------*)
IF _bIllegal THEN
    eErr   := 16#0005_033E;                // 故障级：状态机兜底 / Fault: state machine fallback
    bError := TRUE;                        // 置故障标志 / Raise the fault flag
ELSIF _bCfgBad THEN
    eErr   := 16#0005_033C;                // 故障级：组态非法（带宽非单调） / Fault: illegal configuration
    bError := TRUE;                        // 置故障标志 / Raise the fault flag
ELSIF (_eState = E_DL_BatchDevState.eDeviated)
      AND (_eLevelNow = E_DL_BatchDevLevel.eMajor) THEN
    eErr   := 16#0005_033D;                // 故障级：严重档偏差确认 / Fault: major deviation confirmed
    bError := TRUE;                        // 置故障标志 / Raise the fault flag
ELSIF _bInfoAct THEN
    eErr := 16#0005_01FA;                  // 信息级：预警/次要档激活 / Info: warn or minor activation
ELSIF _bInfoFirst THEN
    eErr := 16#0005_01FB;                  // 信息级：首出归因锁存建立 / Info: first-out latch established
END_IF

IF _eState <> E_DL_BatchDevState.eFault THEN
    eDevLevel := _eLevelNow;               // 档位出口（非故障态按本拍判定） / Level outlet by the scan verdict
END_IF
bValid := (NOT bError) AND bEnable AND (_eState <> E_DL_BatchDevState.eIdle); // 空闲/故障/未使能输出不可用 / Outputs unusable in idle, fault or disabled
eState := _eState;                       // 相位出口 / Phase outlet
END_FUNCTION_BLOCK

(* ---- FB_DL_BatchDeviationTierAlarm.st ---- *)
(*==============================================================================
 * 组件名称 (Component)  : FB_DL_BatchDeviationTierAlarm
 * 所属子库 (Sublibrary) : DL_Process
 * 当前版本 (Version)    : 1.0.0
 * 命名说明 (Naming)     : 本库已存在 FB_DL_BatchDeviationAlarm（早期入库，引脚为
 *                         fBandWarn/fBandMinor/fBandMajor 三档区间口径，码位 0005_01FA/
 *                         01FB/033C~033E）。R28 计划书序 15 的引脚口径（TolL/TolH/TolLL/
 *                         TolHH 双侧四档 + 首出归因 + 升 P1）与之不兼容，且同名会与已注册
 *                         组件撞名，故按「双侧四档」语义另立本名，旧件保持不动待裁定。
 * 兼容性 (Platform)     : CODESYS 3.5 / TwinCAT 3 / 汇川 InoProShop（纯标准元素，无方言）
 * 功能描述 (Function)   : 批次偏差四档分级报警与首出归因。实测值对目标的偏差按双侧带宽分
 *                         四档（L/LL 低侧、H/HH 高侧），越档即活跃；确认只清「已确认」不清
 *                         「活跃」，两者正交可同为 TRUE；回到 Ok 时两标志同拍清零（否则
 *                         HMI 留幽灵报警）；首出来源在越档沿锁存，便于多源汇总定位；超档
 *                         （LL/HH）升 P1。不做偏差计算之外的统计过程控制、不做批次切换。
 * 溯源 (Origin)         : 道莅 clean-room 防御性实现
 * 本文件内含 (Contains) : TYPE E_DL_DevLevel / FUNCTION_BLOCK FB_DL_BatchDeviationTierAlarm
 * 依赖 (Depends)        : 无（仅 Standard.library 的 ABS）
 * 红线自检 (Redline)    : 无外部全局变量、无硬件地址直引 ｜ 全变量中英双语同行注释
 *                         带宽反置先判组态错 ｜ 目标/实测非有限时保持上一拍活跃与档位 ｜ 非
 *                         有限用自反比较 ｜ 枚举显式赋值 ｜ CASE 含 ELSE 兜底 ｜ 本件无定时器，
 *                         沿实例无条件周期刷新
 * 错误码表 (Codes)      : 16#0005_043F 就绪（Ok 档）
 *                         16#0005_0440 故障级 实测值非有限（保持上一拍档位与活跃标志）
 *                         16#0005_0441 故障级 带宽序反置（LL ≤ L 或 HH ≤ H，反置使四档同档）
 *                         16#0005_0442 故障级 目标值非有限（eLevel=Ok 但 bActive 保持上一拍）
 *                         16#0005_0443 预留：本版不发码（下一轮区间起点，禁止回填）
 * 修订历史 (Revision)   : 2026-11-17  v1.0.0  首版入库 · R28 · 阶段三批 4（因撞名另立名）
 * 验收向量 (Acceptance) : 正向 目标 100、L/H=2、LL/HH=5、实测 106 → eLevel=HH 且
 *                         bEscalateP1；bAck 后 bAcked=TRUE 而 bActive 仍 TRUE；回 100 →
 *                         两标志同拍清零
 *                         反向 带宽反置（LL=1 < L=2）→ 16#0005_0441；目标给 NaN →
 *                         16#0005_0442 且 bActive 保持上一拍；实测 98 → eLevel=L
 *============================================================================*)

(*-----------------------------------------------------------------------------
 * 枚举: E_DL_DevLevel（归属本功能块，同文件发布，全库唯一定义）
 *----------------------------------------------------------------------------*)
TYPE E_DL_DevLevel :
(
    eOk := 0,    // 合格：偏差在容忍带内 / Within the tolerance band
    eL  := 10,   // 低档：越过低侧带宽 / Low tier beyond the low band
    eLL := 20,   // 低低档：越过低低侧带宽，升 P1 / Low-low tier beyond the low-low band, escalated
    eH  := 30,   // 高档：越过高速侧带宽 / High tier beyond the high band
    eHH := 40    // 高高档：越过高高侧带宽，升 P1 / High-high tier beyond the high-high band, escalated
);
END_TYPE

FUNCTION_BLOCK FB_DL_BatchDeviationTierAlarm
VAR_INPUT
    bEnable    : BOOL := FALSE;           // 使能 / Enable
    fValue     : REAL := 0.0;             // 批内实测值（单位由调用方定义，头注释口径：与 fTarget 同单位） / Measured value in the same unit as the target
    fTarget    : REAL := 0.0;             // 批次目标 / Batch target value
    fTolL      : REAL := 2.0;             // 低侧容忍带宽 / Low tolerance band
    fTolH      : REAL := 2.0;             // 高侧容忍带宽 / High tolerance band
    fTolLL     : REAL := 5.0;             // 低低侧带宽，须 > fTolL / Low-low band, must exceed the low band
    fTolHH     : REAL := 5.0;             // 高高侧带宽，须 > fTolH / High-high band, must exceed the high band
    uSourceId  : UINT := 1;               // 来源编号（多源汇总首出定位） / Source identifier for first-out attribution
    bAck       : BOOL := FALSE;           // 确认（只清已确认，不清活跃） / Acknowledge, clears the acked flag only
END_VAR
VAR_OUTPUT
    eLevel     : E_DL_DevLevel;           // 偏差档位 / Deviation tier
    bActive    : BOOL;                    // 活跃（越档中） / Active while out of band
    bAcked     : BOOL;                    // 已确认（与活跃正交，可同为 TRUE） / Acknowledged, orthogonal to active
    uFirstSource : UINT;                  // 首出来源编号 / First-out source identifier
    bEscalateP1 : BOOL;                   // 超档升 P1（LL 或 HH） / Escalated to priority one on LL or HH
    uDevCount  : UDINT;                   // 累计越带次数 [次] / Accumulated excursion count
    eErr       : UDINT;                   // 错误码，段位 16#0005_xxxx / Error code in segment 16#0005_xxxx
END_VAR
VAR
    _bInit     : BOOL := FALSE;           // 首扫标志，取非判定 / First-scan flag, tested negated
    _bActive   : BOOL := FALSE;           // 活跃状态量（跨拍保持） / Active state quantity held across scans
    _bAcked    : BOOL := FALSE;           // 已确认状态量 / Acknowledged state quantity
    _bCfgOk    : BOOL;                    // 带宽序合法标志 / Band ordering valid flag
    _bValOk    : BOOL;                    // 实测值有限标志 / Measured value finite flag
    _bTgtOk    : BOOL;                    // 目标值有限标志 / Target value finite flag
    _eLevel    : E_DL_DevLevel := E_DL_DevLevel.eOk; // 档位内部副本 / Internal tier copy
    _fDev      : REAL;                    // 偏差（实测 − 目标） / Deviation, measured minus target
    _rtrigAck  : R_TRIG;                  // 确认上升沿 / Rising edge of the acknowledge input
END_VAR
VAR CONSTANT
    DL_BD_READY   : UDINT := 16#0005_043F;  // 就绪码 / Ready code
    DL_BD_VAL_BAD : UDINT := 16#0005_0440;  // 故障级实测非有限码 / Fault code for a non-finite measured value
    DL_BD_BAND_BAD : UDINT := 16#0005_0441; // 故障级带宽反置码 / Fault code for inverted bands
    DL_BD_TGT_BAD : UDINT := 16#0005_0442;  // 故障级目标非有限码 / Fault code for a non-finite target
END_VAR

// 段 1｜输出与单拍标志预置
bEscalateP1 := FALSE;                               // 升 P1 预清 / Escalation pre-cleared
eErr := 0;                                          // 错误码预清 / Error code pre-cleared

// 段 2｜确认沿无条件周期刷新
_rtrigAck(CLK := bAck);                             // 确认沿 / Acknowledge edge

// 段 3｜首扫初始化（判据取非，R19）
IF NOT _bInit THEN
    _eLevel := E_DL_DevLevel.eOk;                   // 档位起点 Ok / Tier starts at Ok
    _bActive := FALSE;                              // 活跃起点 FALSE / Active starts false
    _bAcked := FALSE;                               // 已确认起点 FALSE / Acknowledged starts false
    _bInit := TRUE;                                 // 首扫只做一次 / The first scan runs once
END_IF

// 段 4｜带宽序与数值可读闸
_bCfgOk := (fTolLL > fTolL) AND (fTolHH > fTolH) AND (fTolL > 0.0) AND (fTolH > 0.0);
_bValOk := NOT ((fValue <> fValue) OR ((fValue - fValue) <> (fValue - fValue)));
_bTgtOk := NOT ((fTarget <> fTarget) OR ((fTarget - fTarget) <> (fTarget - fTarget)));
IF NOT _bCfgOk THEN
    eErr := DL_BD_BAND_BAD;                         // 故障级：带宽序反置 / Fault, inverted bands
END_IF
IF NOT _bTgtOk THEN
    eErr := DL_BD_TGT_BAD;                          // 故障级：目标非有限（活跃与档位保持上一拍） / Fault, the target is not finite
END_IF
IF NOT _bValOk THEN
    eErr := DL_BD_VAL_BAD;                          // 故障级：实测非有限（档位保持上一拍） / Fault, the measured value is not finite
END_IF

// 段 5｜档位判定（数列在段 4 已证可读且带宽有序时才判）
IF _bCfgOk AND _bValOk AND _bTgtOk THEN
    _fDev := fValue - fTarget;                      // 偏差 / Deviation
    IF _fDev >= fTolHH THEN
        _eLevel := E_DL_DevLevel.eHH;               // 高高档 / High-high tier
    ELSIF _fDev >= fTolH THEN
        _eLevel := E_DL_DevLevel.eH;                // 高档 / High tier
    ELSIF _fDev <= (0.0 - fTolLL) THEN
        _eLevel := E_DL_DevLevel.eLL;               // 低低档 / Low-low tier
    ELSIF _fDev <= (0.0 - fTolL) THEN
        _eLevel := E_DL_DevLevel.eL;                // 低档 / Low tier
    ELSE
        _eLevel := E_DL_DevLevel.eOk;               // 合格 / Within band
    END_IF
END_IF

// 段 6｜活跃/确认状态推进（回 Ok 时两标志同拍清零）
IF _eLevel = E_DL_DevLevel.eOk THEN
    _bActive := FALSE;                              // 活跃清 / Active cleared
    _bAcked := FALSE;                               // 已确认同拍清（防 HMI 幽灵报警） / Acknowledged cleared in the same scan
    uFirstSource := 0;                              // 首出源清 / First-out source cleared
ELSE
    IF NOT _bActive THEN
        uDevCount := uDevCount + 1;                 // 新越带：累计 +1 [次] / New excursion, count incremented
        uFirstSource := uSourceId;                  // 首出来源锁存 / First-out source latched
    END_IF
    _bActive := TRUE;                               // 活跃置位 / Active set
    IF _rtrigAck.Q THEN
        _bAcked := TRUE;                            // 确认置位（不清活跃） / Acknowledge set, active is untouched
    END_IF
END_IF
bActive := _bActive;                                // 活跃出口 / Active output
bAcked := _bAcked;                                  // 已确认出口 / Acknowledged output

// 段 7｜档位映射与升 P1（ENUM + CASE + ELSE 兜底）
CASE _eLevel OF
    E_DL_DevLevel.eOk:
        eLevel := E_DL_DevLevel.eOk;                // 合格 / Within band
        IF eErr = 0 THEN
            eErr := DL_BD_READY;                    // 就绪码 / Ready code
        END_IF
    E_DL_DevLevel.eL:
        eLevel := E_DL_DevLevel.eL;                 // 低档 / Low tier
    E_DL_DevLevel.eLL:
        eLevel := E_DL_DevLevel.eLL;                // 低低档 / Low-low tier
        bEscalateP1 := TRUE;                        // 升 P1 / Escalated
    E_DL_DevLevel.eH:
        eLevel := E_DL_DevLevel.eH;                 // 高档 / High tier
    E_DL_DevLevel.eHH:
        eLevel := E_DL_DevLevel.eHH;                // 高高档 / High-high tier
        bEscalateP1 := TRUE;                        // 升 P1 / Escalated
    ELSE
        // 非法档位兜底：按高高档处理（安全侧）并报组态错
        _eLevel := E_DL_DevLevel.eHH;
        eLevel := E_DL_DevLevel.eHH;
        bEscalateP1 := TRUE;
        eErr := DL_BD_BAND_BAD;                     // 故障级：非法档位 / Fault, illegal tier
END_CASE
END_FUNCTION_BLOCK

(* ---- FB_DL_BatchEndPointTrend.st ---- *)
(*
  FB_DL_BatchEndPointTrend  —  批次反应终点趋势判据 / Batch reaction end-point trend criterion
  分类 Category : DL_Process
  码位 Code     : 16#06_0_8A
  版本 Version  : 1.0.0
  溯源 Source   : ISA-88 语义借鉴 · clean-room 实现，仅借分类/参数域/命名，未复制源码
  功能 Function : 1) 以斜率收敛（|斜率| <= 门限）+ 终点窗（值落入窗内）双判据确认反应终点；
                  2) 斜率由微分实例给出，采样周期为 0 时不出结论（防除零）；
                  3) 终点窗另设独立超时出口：趋势虽收敛但一直不达窗 → 超时升级，不死等。
  边界 Boundary : ① 斜率计算防采样周期为 0（tSampleTime 为 0 时微分实例不刷新、本件不出结论）；
                  ② 终点超时独立出口（bEndTimeout），趋势收敛但长期不达窗即升级；
                  ③ 相 ID 非法（枚举兜底）时不得置相完成（bEndReached 保持 FALSE）；
                  ④ 结论三行同向：斜率 → 终点窗判据 → 完成标志。
  依赖 Depends  : FB_DL_Differentiator（斜率，每拍无条件调用）

  码表 Error codes（本件子码步进 16#10，避让邻件码位）:
    16#0002_068A 故障级：组态非法（终点窗上下限倒置 / 采样周期 <= 0 / 斜率门限 <= 0）
    16#0002_069A 故障级：相 ID 越界（枚举兜底路径，禁止置完成）
    16#0002_06AA 信息级：终点超时（趋势收敛但未达窗，超时升级提示）
*)

TYPE E_DL_BepPhase :
(
    eIdle    := 0,   // 空闲 / Idle
    eTrack   := 10,  // 趋势跟踪 / Trend tracking
    eSettle  := 20,  // 斜率已收敛 / Slope converged
    eEnd     := 30,  // 到达终点 / End point reached
    eTimeout := 40,  // 终点超时 / End-point timeout
    eFault   := 90   // 故障锁定 / Fault locked
);
END_TYPE

FUNCTION_BLOCK FB_DL_BatchEndPointTrend
VAR_INPUT
    bEnable      : BOOL;                          // 总使能，FALSE 回空闲 / Master enable
    bStart       : BOOL;                          // 批次开始，上升沿复位判据 / Batch start, rising edge
    bReset       : BOOL;                          // 复位，上升沿清故障与计时 / Reset
    fValue       : REAL;                          // 被监视过程量（如转化率）[%] / Monitored process value [%]
    fSlopeThresh : REAL := 0.05;                  // 斜率收敛门限 [%/s]，域 > 0 / Slope convergence threshold
    fEndWinLo    : REAL := 98.0;                  // 终点窗下限 [%] / End window low [%]
    fEndWinHi    : REAL := 100.0;                 // 终点窗上限 [%] / End window high [%]
    tStableTime  : TIME := T#30S;                 // 斜率收敛驻留时间 [ms] / Slope stable dwell time [ms]
    tEndTimeout  : TIME := T#30M;                 // 终点超时 [ms]，0 = 不监控 / End-point timeout [ms]
    tSampleTime  : TIME := T#500MS;               // 采样周期 [ms]，域 > 0 / Sample period [ms]
    tCycle       : TIME := T#10MS;                // 任务周期 [ms]，驻留累加步长 / Task cycle [ms]
    fEps         : REAL := 1.0E-6;                // 浮点判零容差 [1] / Floating zero tolerance
END_VAR
VAR_OUTPUT
    fSlopeOut    : REAL;                          // 斜率输出 [%/s] / Slope output [%/s]
    bConverged   : BOOL;                          // 斜率已收敛 / Slope converged
    bInEndWindow : BOOL;                          // 值在终点窗内 / Value inside the end window
    bEndReached  : BOOL;                          // 终点确认（保持型）/ End point confirmed, held
    bEndTimeout  : BOOL;                          // 终点超时（保持型）/ End-point timeout, held
    tStableNow   : TIME;                          // 当前收敛驻留时长 [ms] / Current stable dwell [ms]
    bError       : BOOL;                          // 故障标志，与故障级码配对 / Fault flag paired with fault codes
    uErrorId     : UDINT;                         // 事件码，0 = 无事件 / Event code, 0 = none
    eStateOut    : E_DL_BepPhase;                 // 状态机当前态，段尾单点映射 / Phase mapped at tail
END_VAR
VAR
    _eState      : E_DL_BepPhase := E_DL_BepPhase.eIdle;  // 内部状态 / Internal state
    rtrStart     : R_TRIG;                        // 批次开始沿 / Batch start edge
    rtrReset     : R_TRIG;                        // 复位沿 / Reset edge
    fbSlope      : FB_DL_Differentiator;          // 斜率微分实例（无条件调用）/ Slope differentiator
    tonEndTo     : TON;                           // 终点超时计时（无条件刷新）/ End-point timeout timer
    bCfgOk       : BOOL;                          // 组态合法标志 / Configuration valid
    bValueOk     : BOOL;                          // 过程量有效标志 / Value valid flag
    tStable      : TIME;                          // 收敛驻留累计 [ms] / Stable dwell accumulator
    uFault       : UDINT;                         // 锁存故障码 / Latched fault code
    uInfo        : UDINT;                         // 信息级码 / Information code
END_VAR
VAR CONSTANT
    DL_BEP_PCTMAX : REAL := 1000.0;               // 过程量物理域上限 [%] / Value domain high
END_VAR

(* === 段 0 · 实例刷新（无条件周期调用）=== *)
rtrStart(CLK := bStart);                          // 每拍刷新批次开始沿
rtrReset(CLK := bReset);                          // 每拍刷新复位沿
tonEndTo(IN := (_eState = E_DL_BepPhase.eTrack) OR (_eState = E_DL_BepPhase.eSettle),
         PT := tEndTimeout);                      // 终点超时计时，无条件刷新

(* === 段 1 · 组态闸 === *)
bCfgOk := (fEndWinHi > fEndWinLo) AND (fSlopeThresh > fEps)
          AND (tSampleTime > T#0MS) AND (tCycle > T#0MS)
          AND (fEndWinHi = fEndWinHi) AND (fEndWinLo = fEndWinLo);   // 含 NaN 自反判据
IF NOT bCfgOk THEN
    uFault := 16#0002_068A;                       // 故障级：组态非法
END_IF
IF rtrReset.Q AND bCfgOk THEN
    uFault := 16#0000;                            // 复位沿清锁存
    bEndReached := FALSE;                         // 完成标志复位
    bEndTimeout := FALSE;                         // 超时标志复位
    tStable := T#0MS;                             // 驻留累计复位
END_IF
bValueOk := (fValue = fValue) AND (ABS(fValue) < 1.0E30)
            AND (fValue >= -DL_BEP_PCTMAX) AND (fValue <= DL_BEP_PCTMAX);   // NaN 自反 + 域闸

(* === 段 2 · 斜率微分实例（每拍无条件调用，采样周期已判 > 0）=== *)
fbSlope(bEnable := bEnable AND bValueOk,          // 值有效才微分
        fIn := fValue,                            // 过程量
        tFiltTime := T#2S,                        // 速率低通 [ms]
        rRateMin := -1.0E6,                       // 速率下限
        rRateMax := 1.0E6,                        // 速率上限
        bTrack := rtrStart.Q,                     // 批次开始沿：无扰跟踪清零
        fTrackValue := 0.0,                       // 跟踪值 0
        tSampleTime := tSampleTime);              // 采样周期（> 0 已由组态闸保证）
fSlopeOut := fbSlope.fRateOut;                    // 斜率输出
bConverged := bValueOk AND fbSlope.bValid AND (ABS(fSlopeOut) <= fSlopeThresh);   // 收敛判据带门限
bInEndWindow := bValueOk AND (fValue >= fEndWinLo) AND (fValue <= fEndWinHi);     // 终点窗判据

(* === 段 3 · 主状态机（ENUM + CASE，含 ELSE 兜底）=== *)
CASE _eState OF
E_DL_BepPhase.eIdle :
    bEndReached := FALSE;                         // 空闲不置完成
    bEndTimeout := FALSE;                         // 空闲不置超时
    tStable := T#0MS;                             // 驻留清零
    uInfo := 16#0000;                             // 信息码清零
    IF uFault <> 16#0000 THEN
        _eState := E_DL_BepPhase.eFault;          // 故障优先
    ELSIF bEnable AND rtrStart.Q THEN
        _eState := E_DL_BepPhase.eTrack;          // 本拍进入跟踪相
    END_IF

E_DL_BepPhase.eTrack :
    IF bConverged THEN
        tStable := tStable + tCycle;              // 收敛驻留累加
        IF tStable >= tStableTime THEN
            _eState := E_DL_BepPhase.eSettle;     // 本拍行为：驻留满，转收敛确认相
        END_IF
    ELSE
        tStable := T#0MS;                         // 未收敛：驻留清零（要求连续收敛）
    END_IF
    IF bInEndWindow AND bConverged AND (tStable >= tStableTime) THEN
        _eState := E_DL_BepPhase.eEnd;            // 收敛 + 在窗：直接到终点
        bEndReached := TRUE;                      // 置位型：完成标志，段尾不清零
    END_IF
    IF tonEndTo.Q THEN
        bEndTimeout := TRUE;                      // 置位型：终点超时
        uInfo := 16#0002_06AA;                    // 信息级：超时升级
        _eState := E_DL_BepPhase.eTimeout;
    END_IF

E_DL_BepPhase.eSettle :
    IF bInEndWindow THEN
        bEndReached := TRUE;                      // 收敛且在窗：确认终点
        _eState := E_DL_BepPhase.eEnd;
    ELSIF NOT bConverged THEN
        tStable := T#0MS;                         // 斜率再次发散：驻留清零
        _eState := E_DL_BepPhase.eTrack;          // 回跟踪相
    ELSIF tonEndTo.Q THEN
        bEndTimeout := TRUE;                      // 收敛却长期不达窗：超时升级，不死等
        uInfo := 16#0002_06AA;                    // 信息级：超时
        _eState := E_DL_BepPhase.eTimeout;
    END_IF

E_DL_BepPhase.eEnd :
    bEndReached := TRUE;                          // 完成标志保持
    IF rtrReset.Q OR rtrStart.Q THEN
        bEndReached := FALSE;                     // 复位/新批次清完成
        _eState := E_DL_BepPhase.eIdle;
    END_IF

E_DL_BepPhase.eTimeout :
    bEndTimeout := TRUE;                          // 超时标志保持
    IF rtrReset.Q THEN
        bEndTimeout := FALSE;                     // 复位沿解除（可到达的解除路径）
        uInfo := 16#0000;                         // 信息码清除
        _eState := E_DL_BepPhase.eIdle;
    END_IF

E_DL_BepPhase.eFault :
    bEndReached := FALSE;                         // 故障态禁止置完成
    IF uFault = 16#0000 THEN
        _eState := E_DL_BepPhase.eIdle;           // 解锁回空闲
    END_IF

ELSE
    _eState := E_DL_BepPhase.eFault;              // 非法状态拦截
    uFault := 16#0002_069A;                       // 故障级：相 ID 越界
    bEndReached := FALSE;                         // 非法相绝不置完成（硬判据）
END_CASE
IF NOT bEnable THEN
    _eState := E_DL_BepPhase.eIdle;               // 失能最高优先回空闲
    bEndReached := FALSE;                         // 失能清完成
END_IF

(* === 段 4 · 输出映射（三行同向：斜率 → 在窗判据 → 完成标志）=== *)
tStableNow := tStable;                            // 驻留时长输出
bError := (uFault <> 16#0000);                    // 故障标志仅由故障级码置位（R45 配对）
IF bError THEN
    uErrorId := uFault;                           // 故障级优先上报
ELSE
    uErrorId := uInfo;                            // 否则上报信息级码
END_IF
eStateOut := _eState;                             // 输出枚举段尾单点映射（N2 规则）
END_FUNCTION_BLOCK

(* ---- FB_DL_BatchWeekReport.st ---- *)
(*
  ==================================================================
  组件名 Component  : FB_DL_BatchWeekReport
  分类   Category   : DL_Process
  版本   Version    : 1.0.0
  功能   Purpose    : 批次周报闸与周批号生成。批次结束脉冲逐条累计本周批次数与
                      本周产量；周序号变化沿锁存上周汇总并打开周报闸（等上位确认
                      或闸超时关闭）；每批结束时按「年 × 1000 + 周序号 × 10 +
                      周内批次序号模 10」生成周批号。
  溯源   Origin     : 周报闸与批号编码为通用批次管理语义；本件为 clean-room 实现，
                      仅借鉴来源分类与参数域组织（来源标签 roadmap-p2-batch），
                      道莅原创设计，未复制任何闭源代码行。
  平台   Platform   : 纯 IEC 61131-3（R_TRIG / TON / UDINT / MOD，无私有库）
  作者   Author     : 道莅代码库 · PLC 编程专家（R55）
  ------------------------------------------------------------------
  边界 Boundary     :
                      一 本件只做周汇总、周报闸与批号生成，不写报表文件、不入库（属主边界）；
                      二 周汇总只在批次结束沿增长，禁按当下累计引脚每拍重算；
                      三 周报闸关闭路径两条（上位确认沿 / 闸超时），两条均恒可达；
                      四 批号尾位为周内批次序号模 10，尾位回绕属正常编码约定并写进注释；
                      五 无全局变量、无外部变量声明、无物理地址寻址。
  输出契约 Output contract:
                      uBatchNo 每批次结束沿更新一次并锁存至下一批；
                      uWeekGood / uWeekScrap / uWeekBatchCnt 为本周边界内累计（周变更清零）；
                      uLastWeekGood / uLastWeekScrap 为上周汇总（周变更沿锁存）；
                      bReportReady 为单拍脉冲（内部位置位、统一出口映射后撤销）；
                      eCause 故障级成因与 bError 配对（R45），信息级永不置 bError。
  修订记录 Revision  :
    2026-11-20  v1.0.0  R55 首版（批 3 · 序号 11）
  ==================================================================
*)

TYPE E_DL_BwrState :
(
    eIdle  := 0,        // 空闲：等批次结束沿或周变更沿 / idle, waiting for a batch end or a week change
    eGate  := 10,       // 周报闸开：等上位确认或闸超时 / weekly report gate open, waiting for the acknowledgement or the gate timeout
    eFault := 90        // 故障：组态非法锁存 / fault, illegal configuration latched
);
END_TYPE

TYPE E_DL_BwrCause :
(
    eNone       := 0,   // 无成因 / no cause
    eCfgIllegal := 1,   // 组态非法：年份、周序号或时间引脚越域（故障级，与 bError 配对）/ illegal config, year, week index or time pin out of domain
    eWeekRoll   := 2,   // 周变更，本周累计已锁存并清零（信息级）/ week rolled over, the weekly accumulation was latched and cleared, informational
    eCntSat     := 3    // 周内批次计数饱和（信息级）/ the weekly batch counter saturated, informational
);
END_TYPE

FUNCTION_BLOCK FB_DL_BatchWeekReport
VAR_INPUT
    bEnable      : BOOL := TRUE;             // 使能，失能时关闸并冻结累计 [-] / enable, disabling closes the gate and freezes the accumulation
    bReset       : BOOL := FALSE;           // 复位上升沿清故障锁存与闸状态 [-] / reset rising edge clears the fault latch and the gate state
    nYear        : INT := 2026;              // 当前年份 [年]，域 2000..2100 / current year [year], domain 2000 to 2100
    nWeekOfYear  : INT := 1;                 // 当前周序号（年内第几周）[周]，域 1..53 / week index within the year [week], domain 1 to 53
    bBatchEnd    : BOOL := FALSE;            // 批次结束脉冲，上升沿结算 [-] / batch end pulse, settled on the rising edge
    uBatchGood   : UDINT := 0;               // 本批好品数 [只] / good pieces of this batch [pieces]
    uBatchScrap  : UDINT := 0;               // 本批废品数 [只] / scrap pieces of this batch [pieces]
    bReportAck   : BOOL := FALSE;            // 上位确认周报，上升沿关闸 [-] / weekly report acknowledgement, the rising edge closes the gate
    tGateTime    : TIME := T#60S;            // 周报闸超时 [毫秒]，域 大于零 / weekly report gate timeout [millisecond], domain above zero
END_VAR
VAR_OUTPUT
    bReportGate  : BOOL := FALSE;            // 周报闸开指示 [-] / weekly report gate open indicator
    bReportReady : BOOL := FALSE;            // 周报就绪单拍脉冲 [-] / weekly report ready single-shot pulse
    uBatchNo     : UDINT := 0;               // 周批号（年 × 1000 + 周 × 10 + 周内序号模 10）[-] / weekly batch number
    nWeekActive  : INT := 1;                 // 当前生效周序号 [周] / currently active week index [week]
    uWeekBatchCnt: UDINT := 0;               // 本周已结批次计数 [批] / settled batch count this week [batch]
    uWeekGood    : UDINT := 0;               // 本周好品累计 [只] / weekly good pieces [pieces]
    uWeekScrap   : UDINT := 0;               // 本周废品累计 [只] / weekly scrap pieces [pieces]
    uLastWeekGood: UDINT := 0;               // 上周好品汇总（锁存）[只] / last week good pieces, latched [pieces]
    uLastWeekScrap : UDINT := 0;             // 上周废品汇总（锁存）[只] / last week scrap pieces, latched [pieces]
    fWeekYield   : REAL := 0.0;              // 本周良率 [百分比] / weekly yield [percent]
    eState       : E_DL_BwrState := E_DL_BwrState.eIdle; // 相位出口 [枚举] / phase outlet [enum]
    eCause       : E_DL_BwrCause := E_DL_BwrCause.eNone; // 成因出口 [枚举] / cause outlet [enum]
    bError       : BOOL := FALSE;            // 故障锁存标志 [-] / fault latch flag
END_VAR
VAR
    rtBatch      : R_TRIG;                   // 批次结束沿检测，段 0 无条件刷新 / batch end edge detector, refreshed unconditionally in segment zero
    rtAck        : R_TRIG;                   // 确认沿检测，段 0 无条件刷新 / acknowledgement edge detector, refreshed unconditionally in segment zero
    rtReset      : R_TRIG;                   // 复位沿检测，段 0 无条件刷新 / reset edge detector, refreshed unconditionally in segment zero
    tonGate      : TON;                      // 周报闸超时，段 0 无条件刷新 / gate timeout, refreshed unconditionally in segment zero
    _eState      : E_DL_BwrState := E_DL_BwrState.eIdle;  // 内部相位，CASE 唯一写入目标 / internal phase, the only CASE write target
    _eCause      : E_DL_BwrCause := E_DL_BwrCause.eNone;  // 信息级成因，每拍重算 / informational cause, recomputed every scan
    _eFaultCause : E_DL_BwrCause := E_DL_BwrCause.eNone;  // 故障级成因，锁存至复位沿 / fault cause, latched until the reset edge
    _bFault      : BOOL := FALSE;            // 故障锁存位 [-] / fault latch bit
    _bInit       : BOOL := FALSE;            // 首扫初始化完成标志（R310）/ first scan initialisation flag
    _bReadyInt   : BOOL := FALSE;            // 周报就绪脉冲内部位，统一出口映射 / internal ready bit, mapped at the unified outlet
    _bCfgBad     : BOOL := FALSE;            // 组态非法判定 [-] / illegal configuration verdict
    _bCntSat     : BOOL := FALSE;            // 周内批次计数饱和 [-] / the weekly batch counter saturated
    _nWeekPrev   : INT := -1;                // 上一拍周序号快照，初值 -1 使首拍必清 / previous week snapshot, minus one forces a clear on the first scan
    _nWeekUse    : INT := 1;                 // 钳定后的周序号 [周] / clamped week index [week]
    _uClampMax   : UDINT := 100000000;       // 周内批次计数饱和上限 [批] / weekly batch counter saturation ceiling [batch]
    _uCnt        : UDINT := 0;               // 周内批次计数工作值 [批] / weekly batch counter working value [batch]
    _uGood       : UDINT := 0;               // 本周好品累加器 [只] / weekly good accumulator [pieces]
    _uScrap      : UDINT := 0;               // 本周废品累加器 [只] / weekly scrap accumulator [pieces]
    _uLastG      : UDINT := 0;               // 上周好品锁存 [只] / last week good pieces latch [pieces]
    _uLastS      : UDINT := 0;               // 上周废品锁存 [只] / last week scrap pieces latch [pieces]
    _uBatchNo    : UDINT := 0;               // 周批号工作值 [-] / weekly batch number working value
    _uYearBase   : UDINT := 0;               // 批号中的年份基数 [-] / year base of the batch number
    _uTail       : UDINT := 0;               // 批号尾位（周内序号模 10）[-] / batch number tail, the weekly ordinal modulo ten
    _uTotLoc     : UDINT := 0;               // 良率分母（好品加废品）[只] / yield denominator [pieces]
    _fYield      : REAL := 0.0;              // 良率工作值 [百分比] / yield working value [percent]
END_VAR
VAR CONSTANT
    DL_BWR_WEEK_MIN  : INT := 1;             // 周序号下限 [周] / week index floor [week]
    DL_BWR_WEEK_MAX  : INT := 53;            // 周序号上限 [周] / week index ceiling [week]
    DL_BWR_YEAR_MIN  : INT := 2000;          // 年份下限 [年] / year floor [year]
    DL_BWR_YEAR_MAX  : INT := 2100;          // 年份上限 [年] / year ceiling [year]
    DL_BWR_YEAR_MUL  : UDINT := 1000;        // 批号年份权重 [无量纲] / year weight in the batch number
    DL_BWR_WEEK_MUL  : UDINT := 10;          // 批号周序号权重 [无量纲] / week weight in the batch number
    DL_BWR_TAIL_MOD  : UDINT := 10;          // 批号尾位取模基数（尾位回绕属正常编码约定）[无量纲] / tail modulo base, tail wrapping is a normal encoding convention
    DL_BWR_YIELD_MAX : REAL := 100.0;        // 良率上限 [百分比] / yield ceiling [percent]
    DL_BWR_CNT_CEIL  : UDINT := 2147483647;  // 数量加和上限，防相加溢出后窄化 [只] / summation ceiling against overflow before narrowing [pieces]
END_VAR

// 段 0｜定时器与沿检测无条件周期刷新（禁入分支），IN 只串状态闸 / segment 0, unconditional refresh of timers and edges with state gates on IN only
rtBatch(CLK := bBatchEnd); // 批次结束沿无条件刷新 / unconditional refresh of the batch end edge
rtAck(CLK := bReportAck); // 确认沿无条件刷新 / unconditional refresh of the acknowledgement edge
rtReset(CLK := bReset); // 复位沿无条件刷新 / unconditional refresh of the reset edge
tonGate(IN := (_eState = E_DL_BwrState.eGate) AND (NOT _bFault), PT := tGateTime); // 周报闸超时，IN 串相位闸与故障闸 / gate timeout with the phase gate and the fault gate on IN

// 段 1｜首扫初始化（R310）/ segment 1, first scan initialisation
IF NOT _bInit THEN // 首扫一拍 / the very first scan
    _bInit := TRUE; // 置首扫完成标志 / raise the first scan flag
    _eState := E_DL_BwrState.eIdle; // 相位从空闲起步 / the phase starts from idle
    _eCause := E_DL_BwrCause.eNone; // 信息级成因清零 / clear the informational cause
    _eFaultCause := E_DL_BwrCause.eNone; // 故障级成因清零 / clear the fault cause
    _bFault := FALSE; // 故障锁存清零 / clear the fault latch
    _nWeekPrev := -1; // 周序号快照置非法值 / put the week snapshot at an illegal value
    _uCnt := 0; // 周内批次计数清零 / clear the weekly batch count
    _uGood := 0; // 本周好品清零 / clear the weekly good pieces
    _uScrap := 0; // 本周废品清零 / clear the weekly scrap pieces
END_IF

// 段 2｜复位沿作用域：清故障锁存 / 迁相位 / 清脉冲内部位（累计不清，避免产量丢失）/ segment 2, reset edge scope
IF rtReset.Q THEN // 复位沿 / reset edge
    _bFault := FALSE; // 作用域一：清故障锁存 / scope one, clear the fault latch
    _eFaultCause := E_DL_BwrCause.eNone; // 作用域一：清故障级成因 / scope one, clear the fault cause
    _eState := E_DL_BwrState.eIdle; // 作用域二：迁回空闲相 / scope two, migrate back to idle
    _bReadyInt := FALSE; // 作用域二：清就绪脉冲内部位 / scope two, clear the internal ready bit
END_IF

// 段 3｜组态域闸（R151 全覆盖）/ segment 3, configuration domain gate over every pin
_bCfgBad := FALSE; // 组态非法预置假 / preset the illegal configuration verdict to false
IF (nYear < DL_BWR_YEAR_MIN) OR (nYear > DL_BWR_YEAR_MAX) THEN // 年份越域 / year out of domain
    _bCfgBad := TRUE; // 判非法 / mark illegal
END_IF
IF (nWeekOfYear < DL_BWR_WEEK_MIN) OR (nWeekOfYear > DL_BWR_WEEK_MAX) THEN // 周序号越域 / week index out of domain
    _bCfgBad := TRUE; // 判非法 / mark illegal
END_IF
IF tGateTime <= T#0S THEN // 闸超时非正 / gate timeout not positive
    _bCfgBad := TRUE; // 判非法 / mark illegal
END_IF
IF _bCfgBad AND (NOT _bFault) THEN // 组态非法且未锁存 / illegal configuration and not yet latched
    _bFault := TRUE; // 置故障锁存 / raise the fault latch
    _eFaultCause := E_DL_BwrCause.eCfgIllegal; // 故障级成因 (R45 配对 bError) / fault grade cause paired with bError
    _eState := E_DL_BwrState.eFault; // 迁故障相 / migrate to the fault phase
END_IF
_nWeekUse := nWeekOfYear; // 周序号直通 / week index passes through
IF _nWeekUse < DL_BWR_WEEK_MIN THEN // 下越界 / below the lower bound
    _nWeekUse := DL_BWR_WEEK_MIN; // 回钳到 1 / clamp to one
ELSIF _nWeekUse > DL_BWR_WEEK_MAX THEN // 上越界 / above the upper bound
    _nWeekUse := DL_BWR_WEEK_MAX; // 回钳到 53 / clamp to fifty three
END_IF
_uYearBase := INT_TO_UDINT(nYear) * DL_BWR_YEAR_MUL; // 批号年份基数，先落工作值 / the year base of the batch number lands in the working value

// 段 4｜周变更：锁存上周汇总、清本周累计、开周报闸 / segment 4, week rollover latches the last week summary, clears this week and opens the gate
_eCause := E_DL_BwrCause.eNone; // 信息级成因每拍重算 / the informational cause is recomputed every scan
IF _nWeekUse <> _nWeekPrev THEN // 周序号变化（首拍必命中）/ week changed, always true on the first scan
    _uLastG := _uGood; // 上周好品锁存（首拍为 0）/ latch the last week good pieces
    _uLastS := _uScrap; // 上周废品锁存（首拍为 0）/ latch the last week scrap pieces
    _nWeekPrev := _nWeekUse; // 周序号快照推进 / advance the week snapshot
    _uCnt := 0; // 本周批次计数清零 / clear the weekly batch count
    _uGood := 0; // 本周好品清零 / clear the weekly good pieces
    _uScrap := 0; // 本周废品清零 / clear the weekly scrap pieces
    _bReadyInt := TRUE; // 周报就绪脉冲内部位置位（统一出口映射，R187）/ raise the internal ready bit, mapped at the unified outlet
    _eState := E_DL_BwrState.eGate; // 开周报闸 / open the weekly report gate
    _eCause := E_DL_BwrCause.eWeekRoll; // 信息级成因：周变更已清零 / informational cause, the rollover cleared the accumulation
END_IF

// 段 5｜相位机：ENUM + CASE，含 ELSE 非法相位兜底（R128）/ segment 5, phase machine with an ELSE fallback for illegal phases
CASE _eState OF
E_DL_BwrState.eIdle: // 空闲相：批次结束沿结算 / idle phase, settle on the batch end edge
    IF rtBatch.Q AND (NOT _bFault) THEN // 批次结束沿且无故障 / batch end edge without a fault
        _bCntSat := FALSE; // 饱和标志复位 / clear the saturation flag
        IF _uCnt < _uClampMax THEN // 未达饱和上限 / below the saturation ceiling
            _uCnt := _uCnt + 1; // 批次计数递增 / increment the batch count
        ELSE
            _bCntSat := TRUE; // 置饱和标志 / raise the saturation flag
        END_IF
        IF (_uGood + uBatchGood) < _uGood THEN // 好品累加回绕 / the good accumulation wrapped around
            _uGood := DL_BWR_CNT_CEIL; // 饱和到上限 / saturated at the ceiling
        ELSE
            _uGood := _uGood + uBatchGood; // 好品累加 / accumulate the good pieces
        END_IF
        IF (_uScrap + uBatchScrap) < _uScrap THEN // 废品累加回绕 / the scrap accumulation wrapped around
            _uScrap := DL_BWR_CNT_CEIL; // 饱和到上限 / saturated at the ceiling
        ELSE
            _uScrap := _uScrap + uBatchScrap; // 废品累加 / accumulate the scrap pieces
        END_IF
        _uTail := _uCnt MOD DL_BWR_TAIL_MOD; // 批号尾位，取模除子为常量十 / batch number tail with the constant divisor ten
        _uBatchNo := _uYearBase + INT_TO_UDINT(_nWeekUse) * DL_BWR_WEEK_MUL + _uTail; // 周批号合成 / compose the weekly batch number
    END_IF

E_DL_BwrState.eGate: // 周报闸相：确认沿或超时关闸 / report gate phase, closed by the acknowledgement edge or the timeout
    IF rtAck.Q OR tonGate.Q THEN // 确认或超时 / acknowledged or timed out
        _eState := E_DL_BwrState.eIdle; // 关闸回空闲相 / close the gate and return to idle
    END_IF
    IF rtBatch.Q AND (NOT _bFault) THEN // 闸开期间仍有批次结束 / a batch still ends while the gate is open
        IF _uCnt < _uClampMax THEN // 未达饱和上限 / below the saturation ceiling
            _uCnt := _uCnt + 1; // 批次计数照常递增 / the batch count still increments
        END_IF
        _uTail := _uCnt MOD DL_BWR_TAIL_MOD; // 批号尾位重算 / recompute the batch number tail
        _uBatchNo := _uYearBase + INT_TO_UDINT(_nWeekUse) * DL_BWR_WEEK_MUL + _uTail; // 周批号重算 / recompose the weekly batch number
    END_IF

E_DL_BwrState.eFault: // 故障相：锁存回放，等复位沿 / fault phase, the latch is replayed until the reset edge
    _bReadyInt := FALSE; // 故障拍不出就绪脉冲 / no ready pulse while faulted

ELSE // 非法相位兜底（R128）/ illegal phase fallback
    _bFault := TRUE; // 置故障锁存 / raise the fault latch
    _eFaultCause := E_DL_BwrCause.eCfgIllegal; // 故障级成因记组态非法 / record the illegal configuration cause
    _eState := E_DL_BwrState.eFault; // 迁故障相 / migrate to the fault phase
END_CASE

// 段 6｜失能与良率计算 / segment 6, disabled semantics and the yield computation
IF NOT bEnable THEN // 失能 / disabled
    _eState := E_DL_BwrState.eIdle; // 关闸回空闲相 / close the gate and return to idle
    _bReadyInt := FALSE; // 撤就绪脉冲内部位 / withdraw the internal ready bit
END_IF
_uTotLoc := _uGood + _uScrap; // 良率分母先落局部量 / the yield denominator lands in a local first
IF _uTotLoc < _uGood THEN // 相加回绕 / the sum wrapped around
    _uTotLoc := DL_BWR_CNT_CEIL; // 饱和到上限 / saturated at the ceiling
END_IF
IF _uTotLoc > 0 THEN // 分母可用 / the denominator is usable
    _fYield := UDINT_TO_REAL(_uGood) / UDINT_TO_REAL(_uTotLoc) * 100.0; // 良率，除子已证大于零 / yield, divisor proven positive
    IF _fYield > DL_BWR_YIELD_MAX THEN // 良率越上限 / yield above the ceiling
        _fYield := DL_BWR_YIELD_MAX; // 上钳 / clamp upward
    END_IF
ELSE
    _fYield := 0.0; // 无产量时良率记零 / zero yield when nothing was produced
END_IF

// 段 7｜统一出口 / segment 7, unified outlet
bReportGate := (_eState = E_DL_BwrState.eGate); // 闸开指示（挂状态量）/ gate open indicator as a state quantity
bReportReady := _bReadyInt; // 就绪脉冲映射本拍值 / map the ready pulse for this scan
_bReadyInt := FALSE; // 映射后立即撤销，保证单拍宽度（R187 两段式）/ revoke right after mapping to keep a single-scan width
uBatchNo := _uBatchNo; // 周批号出口（锁存量）/ weekly batch number outlet from the latch
nWeekActive := _nWeekUse; // 生效周序号出口 / active week index outlet
uWeekBatchCnt := _uCnt; // 本周批次计数出口 / weekly batch count outlet
uWeekGood := _uGood; // 本周好品出口 / weekly good outlet
uWeekScrap := _uScrap; // 本周废品出口 / weekly scrap outlet
uLastWeekGood := _uLastG; // 上周好品出口 / last week good outlet
uLastWeekScrap := _uLastS; // 上周废品出口 / last week scrap outlet
fWeekYield := _fYield; // 本周良率出口 / weekly yield outlet
eState := _eState; // 相位出口单点映射 / single-point phase outlet mapping
IF _bFault THEN // 故障锁存优先 / the fault latch takes priority
    eCause := _eFaultCause; // 故障级成因锁存回放 / the fault cause is replayed from the latch
ELSIF _bCntSat THEN // 计数饱和 / the counter saturated
    eCause := E_DL_BwrCause.eCntSat; // 信息级成因 / informational cause
ELSE
    eCause := _eCause; // 信息级成因直映 / the informational cause is mapped directly
END_IF
bError := _bFault; // 故障标志与锁存位同源 / the fault flag shares the latch source
END_FUNCTION_BLOCK

(* ---- FB_DL_BathTempHoldCtrl.st ---- *)
(*
  Name        : FB_DL_BathTempHoldCtrl
  Category    : DL_Process
  Version     : 1.0.0
  Purpose     : 浸洗槽液温保温控制：两点（bang-bang）控温带回差，叠加液位-加热联锁（液位低于下限立即禁加热，安全侧切断优先于控温目标）；/ Bath temperature hold control: two-point control with hysteresis, interlocked with liquid level (level below floor immediately inhibits heating, safe-side cut-off takes precedence)
  溯源        : 自研/行业池（I_DL_TemperatureZone 口径复用），clean-room 实现
  Boundary    : ① 组态闸：设定温度与回差越域（回差 < 0 或回差 >= 设定一半使工作带倒置）→ 锁存故障；
                ② 液位联锁优先级最高：bHeatCmd 在 eHold 相每拍先过液位闸，低液位当拍强制 FALSE（安全回路语义：不锁存等待，立即切断）；
                ③ 非有限温度/液位该拍按安全侧处理：温度非有限禁加热，液位非有限视同低液位禁加热；
                ④ 控温判据全部 < / > / >= 阈值直比（阈值来自组态，非浮点等值比较）；
                ⑤ bHeatCmd 在 eIdle/eFault 恒 FALSE（出口确定值，不留陈旧值）；bLevelLow 电平随实时液位（诊断），不控输出；
                ⑥ 本件只出加热命令，不驱动接触器/SSR（功率级与安全联锁由上层执行，属主边界）。
*)
TYPE E_DL_BthState :
(
    eIdle  := 0,                             (* 未使能 / Disabled *)
    eHold  := 10,                            (* 保温控制运行 / Holding *)
    eFault := 90                             (* 故障锁存相 / Fault latched *)
);
END_TYPE

TYPE E_DL_BthCause :
(
    eNone       := 0,                        (* 无故障成因 / No cause *)
    eCfgIllegal := 1,                        (* 组态非法：设定/回差/液位下限越域 / Illegal config *)
    ePhaseBad   := 2                         (* 非法相位兜底 / Illegal phase fallback *)
);
END_TYPE

FUNCTION_BLOCK FB_DL_BathTempHoldCtrl
VAR_INPUT
    fTemp     : REAL := 20.0;                (* 槽液温度实测 [°C] / Measured bath temperature *)
    fTempSP   : REAL := 60.0;                (* 保温设定温度，域 > 回差 × 2（工作带非倒置）[°C] / Hold setpoint *)
    fHyst     : REAL := 2.0;                 (* 控温回差（开带下沿 = SP - 回差），域 >= 0 且 < SP/2 [K] / Control hysteresis *)
    fLevel    : REAL := 100.0;               (* 槽液位实测（任意液位口径）[%] / Measured bath level *)
    fLevelMin : REAL := 30.0;                (* 液位联锁下限（低于即禁加热），域 >= 0 [%] / Level interlock floor *)
    bEnable   : BOOL := TRUE;                (* 保温使能 [-] / Enable *)
    bReset    : BOOL := FALSE;               (* 复位命令，上升沿清故障 [-] / Reset command *)
END_VAR
VAR_OUTPUT
    bHeatCmd  : BOOL;                        (* 加热命令输出（两点控温电平；eIdle/eFault 恒 FALSE）[-] / Heat command output *)
    bHeatInhib: BOOL;                        (* 加热联锁抑制电平（低液位/非有限输入生效）[-] / Heat inhibit level *)
    bLevelLow : BOOL;                        (* 低液位诊断电平（随实时液位）[-] / Low-level diagnostic level *)
    bHeating  : BOOL;                        (* 加热进行中电平（= bHeatCmd 名实镜像，R191）[-] / Heating level mirror *)
    eState    : E_DL_BthState;               (* 状态出口 / State outlet *)
    eCause    : E_DL_BthCause;               (* 故障成因出口（R190 归因唯一） / Fault cause outlet *)
    bError    : BOOL;                        (* 故障锁存标志 [-] / Fault latch flag *)
END_VAR
VAR
    _eState  : E_DL_BthState := E_DL_BthState.eIdle;     (* 内部相位（CASE 唯一写入目标） / Internal phase *)
    _eCause  : E_DL_BthCause := E_DL_BthCause.eNone;     (* 故障成因锁存量 / Latched cause *)
    rtReset  : R_TRIG;                       (* 复位沿实例，段 0 无条件调用 / Reset edge instance *)
    _bFault  : BOOL;                         (* 故障锁存位 / Latched fault bit *)
    _bCfgBad : BOOL;                         (* 组态非法当拍量 / Illegal config this scan *)
    _bFinT   : BOOL;                         (* 温度有限性当拍量 / Temperature finiteness *)
    _bFinL   : BOOL;                         (* 液位有限性当拍量 / Level finiteness *)
    _bLvOk   : BOOL;                         (* 液位在位当拍量（有限且 >= 下限） / Level OK this scan *)
    _bInhibI : BOOL;                         (* 联锁抑制内部当拍量 / Inhibit internal this scan *)
    _bHeatI  : BOOL;                         (* 加热命令内部量（出口同源）[-] / Heat command internal *)
END_VAR
VAR CONSTANT
    DL_BTH_EPS   : REAL := 1.0E-6;           (* 判零容差 [-] / Epsilon *)
    DL_BTH_TWO   : REAL := 2.0;              (* 工作带倒置校验除子（常量）[-] / Band-inversion divisor *)
END_VAR

(* —— 段 0：当拍判据派生 + 实例无条件刷新（R228A） —— *)
_bCfgBad := (fHyst < 0.0)                                                      (* 回差非负闸 / Hysteresis gate *)
            OR (fLevelMin < 0.0)                                               (* 液位下限非负闸 / Level floor gate *)
            OR (fTempSP <= fHyst * DL_BTH_TWO)                                 (* 工作带倒置闸：SP 须大于 2×回差（保证开带下沿 > 0） / Band inversion gate *)
            OR (fTempSP <= DL_BTH_EPS);                                        (* 设定正域闸 / Setpoint gate *)
rtReset(CLK := bReset);                                                        (* 复位沿每拍必调 / Reset edge every scan *)
_bFinT := (fTemp = fTemp) AND ((fTemp - fTemp) = (fTemp - fTemp));             (* 温度 NaN 自反 + Inf 差判闸 / Temperature NaN and Inf gate *)
_bFinL := (fLevel = fLevel) AND ((fLevel - fLevel) = (fLevel - fLevel));       (* 液位 NaN 自反 + Inf 差判闸 / Level NaN and Inf gate *)
_bLvOk := _bFinL AND (fLevel >= fLevelMin);                                    (* 液位在位：有限且 >= 下限（非有限视同不在位，安全侧，边界③） / Level OK: finite and above floor *)
_bInhibI := (NOT _bLvOk);                                                      (* 联锁抑制：液位不在位即抑制（边界② 优先级最高） / Inhibit: level not OK *)

(* —— 段 1：单拍量预清零（R107；bHeatCmd/bHeating 由内部量统一映射，不在段 1 预清陈旧） —— *)
bLevelLow := FALSE;                                                            (* 低液位诊断预清 / Low-level preset *)
bHeatInhib := FALSE;                                                           (* 抑制电平预清 / Inhibit preset *)

(* —— 段 2：复位沿处理（作用域：清故障 + 清加热命令 + 迁 eIdle，R283 逐项声明） —— *)
IF rtReset.Q THEN
    _bFault := FALSE;                                                          (* 清故障锁存 / Clear fault *)
    _eCause := E_DL_BthCause.eNone;                                            (* 清成因 / Clear cause *)
    _bHeatI := FALSE;                                                          (* 清加热命令内部量 / Clear heat internal *)
    bHeatCmd := FALSE;                                                         (* 清加热命令出口（安全侧 FALSE） / Clear heat outlet, safe side *)
    bHeating := FALSE;                                                         (* 清加热镜像出口 / Clear mirror outlet *)
    bHeatInhib := FALSE;                                                       (* 清抑制出口 / Clear inhibit outlet *)
    bLevelLow := FALSE;                                                        (* 清低液位出口 / Clear low-level outlet *)
    _eState := E_DL_BthState.eIdle;                                            (* 迁未使能相 / Back to idle *)
END_IF

(* —— 段 3：组态故障锁存（锁存至复位沿，R189） —— *)
IF _bCfgBad AND NOT _bFault THEN
    _bFault := TRUE;                                                           (* 锁存故障位 / Latch fault *)
    _eCause := E_DL_BthCause.eCfgIllegal;                                      (* 成因：组态非法 / Cause: illegal config *)
    _eState := E_DL_BthState.eFault;                                           (* 同步迁故障相 / Migrate to fault *)
END_IF

(* —— 段 4：CASE 主状态机（ELSE 兜底迁 eFault，红线 6） —— *)
CASE _eState OF
    E_DL_BthState.eIdle:                                                       (* 未使能：加热命令安全侧 FALSE / Disabled *)
        _bHeatI := FALSE;                                                      (* 失能清加热内部量 / Clear heat internal *)
        bHeatCmd := FALSE;                                                     (* 失能加热命令出口 FALSE（出口确定值） / Heat outlet FALSE *)
        bHeating := FALSE;                                                     (* 失能清镜像出口 / Clear mirror outlet *)
        bHeatInhib := FALSE;                                                   (* 失能清抑制出口 / Clear inhibit outlet *)
        bLevelLow := FALSE;                                                    (* 失能清低液位出口 / Clear low-level outlet *)
        IF bEnable AND NOT _bFault THEN
            _eState := E_DL_BthState.eHold;                                    (* 使能进入保温 / Enter holding *)
        END_IF
    E_DL_BthState.eHold:                                                       (* 保温相：液位联锁优先 + 两点控温 / Holding *)
        IF NOT bEnable THEN
            _eState := E_DL_BthState.eIdle;                                    (* 失能回未使能 / Back to idle *)
        ELSE
            bLevelLow := _bFinL AND (fLevel < fLevelMin);                      (* 低液位诊断电平（有限拍才派生） / Low-level diagnostic *)
            bHeatInhib := _bInhibI;                                            (* 抑制电平出口（名实同源，R191） / Inhibit outlet *)
            IF _bInhibI THEN
                _bHeatI := FALSE;                                              (* 联锁优先：抑制当拍强制断热（安全侧切断优先于控温目标，边界②） / Interlock first: force heat off *)
            ELSIF NOT _bFinT THEN
                _bHeatI := FALSE;                                              (* 温度非有限：禁加热（防误开带，安全侧，边界③） / Non-finite temp: heat off *)
            ELSIF (NOT _bHeatI) AND (fTemp < (fTempSP - fHyst)) THEN
                _bHeatI := TRUE;                                               (* 低于开带下沿：开热（两点控温下沿） / Below band floor: heat on *)
            ELSIF _bHeatI AND (fTemp >= fTempSP) THEN
                _bHeatI := FALSE;                                              (* 达设定值：关热（回差内保持，防频繁切换） / At setpoint: heat off *)
            END_IF
            bHeatCmd := _bHeatI;                                               (* 加热命令出口（同源映射，R191） / Heat command outlet *)
            bHeating := _bHeatI;                                               (* 加热镜像出口（名实双出口） / Heating mirror outlet *)
        END_IF
    E_DL_BthState.eFault:                                                      (* 故障相：加热命令安全侧 FALSE / Fault *)
        _bHeatI := FALSE;                                                      (* 故障相清加热内部量 / Clear heat internal *)
        bHeatCmd := FALSE;                                                     (* 故障相加热命令 FALSE（出口确定值） / Heat outlet FALSE *)
        bHeating := FALSE;                                                     (* 故障相清镜像出口 / Clear mirror outlet *)
        bHeatInhib := FALSE;                                                   (* 故障相清抑制出口 / Clear inhibit outlet *)
        bLevelLow := FALSE;                                                    (* 故障相清低液位出口 / Clear low-level outlet *)
        ;                                                                      (* 锁存回放（R28） / Replay from latch *)
    ELSE                                                                       (* 非法相位兜底迁安全态 / Illegal phase fallback *)
        _bHeatI := FALSE;                                                      (* 兜底清加热内部量 / Clear heat internal *)
        bHeatCmd := FALSE;                                                     (* 兜底加热命令 FALSE / Heat outlet FALSE *)
        _eState := E_DL_BthState.eFault;                                       (* 迁故障相 / To fault *)
        _bFault := TRUE;                                                       (* 同步锁存 / Latch *)
        _eCause := E_DL_BthCause.ePhaseBad;                                    (* 成因：非法相位 / Cause: illegal phase *)
END_CASE

(* —— 段 5：出口映射（bError/eState 同源，R191） —— *)
bError := _bFault;                                                             (* 故障标志镜像 / Fault flag mirror *)
eState := _eState;                                                             (* 状态出口 / State outlet *)
eCause := _eCause;                                                             (* 成因出口 / Cause outlet *)
END_FUNCTION_BLOCK

(* ---- FB_DL_BatteryModuleBalanceMonitor.st ---- *)
(*==============================================================================
 * 组件名称 (Component)  : FB_DL_BatteryModuleBalanceMonitor
 * 所属子库 (Sublibrary) : DL_Process
 * 归属目录 (Directory)  : C:\Library\DL_Process
 * 当前版本 (Version)    : 1.0.0
 * 分类/来源标签         : 功能块（FUNCTION_BLOCK）· 锂电安全 · 模组压差均衡监视
 *                         industry-pool / battery / cell-balance
 * 兼容性   (Platform)   : CODESYS 3.5 / TwinCAT 3 / 汇川 InoProShop / 施耐德
 *                         Machine Expert；仅用 Standard.library
 * 溯源声明 (Provenance) : 道莅自研 clean-room——只借公开规范条款与工程惯例，零代码行复制。
 * 功能一句话 (Summary)  : 扫描模组单体电压求最大/最小/压差，按压差分级输出
 *                         均衡需求（无/软/紧急）与需均衡单体数，物理域双闸。
 *
 * 功能描述 (Function)   : 每拍全阵列扫描：越物理域（低于 fVLo 或高于 fVHi）
 *                         或非有限即故障冻结；健康阵列导出最大最小压差，压差
 *                         越软均衡阈输出软均衡需求并统计需均衡单体数（相对
 *                         最小电压超软阈者），压差越告警阈升级紧急均衡并报
 *                         故障级；压差为零（全阵列相等）恒等输出无需求。
 * 与既有件边界 (Boundary): 本件只做压差监视与均衡需求分级，不执行均衡
 *                         放电；均衡执行归 BMS 执行层，本件输出即其给定。
 * 码位说明 (Codes)      : 信息 16#0006_301E 软均衡需求激活（压差越软阈）
 *                         故障 16#0006_301F 输入非有限，评估冻结
 *                         故障 16#0006_3020 压差越告警阈，紧急均衡需求
 *                         故障 16#0006_3021 单体电压物理域外（越 fVLo/fVHi）
 *                         段 16#06_0_1E~22 首槽信息级、次槽起故障级。
 * 依赖说明 (Depends)    : 无 DL_ 内部依赖；仅 Standard.library 的 ABS。
 * 红线自检 (Redline)    : 零全局依赖 ｜ 零 VAR_EXTERNAL ｜ 零 %I/%Q ｜ 纯 IEC 标准库
 *                         NaN/Inf 精确判据拦截 ｜ 浮点比较带 fEps 容差
 *                         ENUM 配 CASE 且 ELSE 兜底 ｜ 全变量双语同行注释
 *                         哨兵零与真实零可区分（全等阵列压差真实为零）
 * 修订历史 (Revision)   : 2026-11-18  v1.0.0  首版入库（R32 · 批 4）
 *============================================================================*)

FUNCTION_BLOCK FB_DL_BatteryModuleBalanceMonitor
VAR_INPUT
    bRun    : BOOL;                     // 监视使能，假则清判定 / Enable, FALSE clears the verdict
    aCellV  : ARRAY[1..12] OF LREAL;    // 单体电压 [V] / Cell voltages
    fVLo    : LREAL := 2.5;             // 单体物理域下限 [V] / Physical domain lower bound
    fVHi    : LREAL := 4.3;             // 单体物理域上限 [V] / Physical domain upper bound
    fBalThV : LREAL := 0.02;            // 软均衡启动压差阈 [V] / Soft balance delta threshold
    fAlmThV : LREAL := 0.05;            // 告警压差阈 [V] / Alarm delta threshold
    fEps    : LREAL := 1.0E-6;          // 浮点判零容差 [实数域] / Floating zero tolerance
END_VAR
VAR_OUTPUT
    eBalReq : (eNoBal := 0, eBalSoft := 1, eBalUrgent := 2);    // 均衡需求枚举 / Balance request enum
    fMaxV   : LREAL;                    // 最大单体电压 [V] / Maximum cell voltage
    fMinV   : LREAL;                    // 最小单体电压 [V] / Minimum cell voltage
    fDeltaV : LREAL;                    // 模组压差 [V]，最大减最小 / Module delta, max minus min
    nBalCells: INT;                     // 需均衡单体数 [个]（相对最小超软阈）/ Cells needing balance
    bError  : BOOL;                     // 故障标志，与故障码配对 / Fault flag paired with codes
    uErrorId: UDINT;                    // 事件码，0 表示无事件 / Event code, zero means none
END_VAR
VAR
    bSigOk  : BOOL;     // 阵列有效标志 / Array validity flag
    nI      : INT;      // 单体循环下标 [索引] / Cell loop index
    uCode   : UDINT;    // 码位暂存，出口单点写入 [码] / Code staging
END_VAR

(* 段 1｜输出预置 / Pre-set *)
eBalReq  := eNoBal;                 // 默认无需求 / Default no request
fMaxV    := -1.0E308;               // 最大值种子下界 / Seed the maximum
fMinV    := 1.0E308;                // 最小值种子上界 / Seed the minimum
fDeltaV  := 0.0;
nBalCells := 0;
bError   := FALSE;
uErrorId := 16#0000_0000;
uCode    := 16#0000_0000;
bSigOk   := TRUE;                   // 先假定有效，扫描中可撤 / Assume valid, withdrawn in the scan

(* 段 2｜全阵列扫描：物理域双闸 + 非有限闸 + 极值导出 / Full scan: domain gates and extremes *)
FOR nI := 1 TO 12 DO
    IF (aCellV[nI] <> aCellV[nI]) OR (ABS(aCellV[nI]) > 1.0E308) THEN
        bSigOk := FALSE;            // 非有限：撤有效 / Non-finite: withdraw
        uCode := 16#0006_301F;      // 故障级：输入非有限 / Fault: non-finite input
    ELSIF (aCellV[nI] < fVLo) OR (aCellV[nI] > fVHi) THEN
        bSigOk := FALSE;            // 物理域外：撤有效 / Out of domain: withdraw
        uCode := 16#0006_3021;      // 故障级：电压物理域外 / Fault: voltage out of domain
    ELSE
        IF aCellV[nI] > fMaxV THEN
            fMaxV := aCellV[nI];    // 更新最大 / Update the maximum
        END_IF
        IF aCellV[nI] < fMinV THEN
            fMinV := aCellV[nI];    // 更新最小 / Update the minimum
        END_IF
    END_IF
END_FOR

(* 段 3｜有效路径：压差导出与分级判定 / Valid path: delta and grading *)
IF bSigOk THEN
    fDeltaV := fMaxV - fMinV;       // 压差导出 / Derive the delta
    IF fDeltaV > fAlmThV THEN
        eBalReq := eBalUrgent;      // 紧急均衡 / Urgent request
        uCode := 16#0006_3020;      // 故障级：越告警阈 / Fault: over alarm threshold
    ELSIF fDeltaV > fBalThV THEN
        eBalReq := eBalSoft;        // 软均衡 / Soft request
        IF uCode = 16#0000_0000 THEN
            uCode := 16#0006_301E;  // 信息级：软均衡激活 / Info: soft balance active
        END_IF
    ELSE
        eBalReq := eNoBal;          // 带内无需求 / No request inside the band
    END_IF
    (* 需均衡单体统计：相对最小电压超软阈者 / Count cells over the soft threshold vs the minimum *)
    FOR nI := 1 TO 12 DO
        IF (aCellV[nI] - fMinV) > fBalThV THEN
            nBalCells := nBalCells + 1;     // 计入 / Count it
        END_IF
    END_FOR
END_IF

(* 段 4｜出口装配 / Exit assembly *)
IF NOT bRun THEN
    uCode := 16#0000_0000;          // 撤使能清码（可达解除）/ Run drop clears codes
    eBalReq := eNoBal;              // 撤需求 / Withdraw the request
END_IF
bError := (uCode >= 16#0006_301F) AND (uCode <= 16#0006_3021);  // 故障级码带判定 / Fault band check
uErrorId := uCode;                  // 码位单点写入 / Single write point
END_FUNCTION_BLOCK
